// TwinCAT 3 PLC project IAG50cmTests
// Title: IAG50cmTests
// Company: BROT
// ProjectVersion: 0.1.0
// ProgramVersion: 3.1.4024.66
// libraries:
//   AstroBROT, 0.5.0 (BROT)
//   BROTLib, 0.20.0 (BROT)
//   Tc2_Math, * (Beckhoff Automation GmbH)
//   Tc3_MC2_AdvancedHoming, * (Beckhoff Automation GmbH)
//   Tc2_MC2, * (Beckhoff Automation GmbH)
//   Tc2_MC2_Drive, * (Beckhoff Automation GmbH)
//   Tc2_NC, * (Beckhoff Automation GmbH)
//   Tc2_Standard, * (Beckhoff Automation GmbH)
//   Tc2_System, * (Beckhoff Automation GmbH)
//   Tc2_Utilities, * (Beckhoff Automation GmbH)
//   Tc3_Module, * (Beckhoff Automation GmbH)
//   TcUnit, * (www.tcunit.org)
// project tree:
//   / PlcTask.TcTTO
//   POUs/ FB_HomeDropReason_Tests.TcPOU, FB_HomeHold_Tests.TcPOU, FB_SweepStop_Tests.TcPOU, FB_PointingModelForward_Tests.TcPOU, FB_TelescopeControl.TcPOU (not stored), FB_HourAngleControl.TcPOU (not stored), FB_DeclinationControl.TcPOU (not stored), FB_AxisControl.TcPOU (not stored), FB_LatchHome.TcPOU (not stored), FB_CabinetControl.TcPOU (not stored), FB_PointingModelInversion.TcPOU (not stored), F_HourAngleOffsetOnAxis.TcPOU (not stored), F_RoundLREAL.TcPOU (not stored), NCError_TO_STRING.TcPOU (not stored), ST_AxisStatus.TcDUT (not stored), FB_AxisMockCore.TcPOU, FB_HourAngleMock.TcPOU, FB_DeclinationMock.TcPOU, FB_FocusMock.TcPOU, FB_CoversMock.TcPOU, FB_DomeMock.TcPOU, FB_NullComm.TcPOU, FB_IagRig_Tests.TcPOU, FB_IagRig.TcPOU, IagStopDuringSlew_Tests.TcPOU, IagCommandInputs_Tests.TcPOU, IagCommandAcceptance_Tests.TcPOU, IagAbortStop_Tests.TcPOU, IagParkPowerReset_Tests.TcPOU, IagSupersede_Tests.TcPOU, IagStuckStop_Tests.TcPOU, GVL_Diag.TcGVL, F_Note.TcPOU, IagResetUnderMotion_Tests.TcPOU, IagTimeouts_Tests.TcPOU, IagErrorPark_Tests.TcPOU, IagParkDuringPowerOn_Tests.TcPOU, IagStopDuringPark_Tests.TcPOU, IagParkInLimit_Tests.TcPOU, FB_RecordingComm.TcPOU, F_NoteNear.TcPOU, FB_IagCoordinatesLegacy.TcPOU, IagTelemetry_Tests.TcPOU, IagCoordinates_Tests.TcPOU, MAIN.TcPOU, FB_HomeDropReason.TcPOU (not stored), FB_HomeHold.TcPOU (not stored), FB_StartRequest.TcPOU (not stored), FB_StartRequest_Tests.TcPOU, FB_StepDrain.TcPOU (not stored), FB_StepDrain_Tests.TcPOU, FB_SweepStop.TcPOU (not stored), FB_PointingModelForward.TcPOU (not stored), GVL_Homing.TcGVL (not stored), GVL_Pointing.TcGVL (not stored)
// real-time tasks:
//   TASK PlcTask: cycle T#10ms, priority 20, ADS port 350

CONFIGURATION IAG50cmTests
    RESOURCE PLC ON TwinCAT3
        TASK PlcTask(INTERVAL := T#10ms, PRIORITY := 20);
        PROGRAM MAIN WITH PlcTask : MAIN;
    END_RESOURCE
END_CONFIGURATION

// ---- POUs/GVL_Diag.TcGVL
{attribute 'qualified_only'}
VAR_GLOBAL
	// the failed checks of the scenario tests (F_Note), one "test: message;" each. Run-Tests.ps1 prints it when a test failed:
	// TcUnit itself only writes the failure text to the ADS log, which CI cannot see.
	sFailures	: STRING(1000);
END_VAR

// ---- POUs/MAIN.TcPOU
PROGRAM MAIN
VAR
	// TcUnit finds every FB_TestSuite instance by itself; it is enough to declare them here.
	fbHomeDropReasonTests	: FB_HomeDropReason_Tests;
	fbHomeHoldTests			: FB_HomeHold_Tests;
	fbStartRequestTests		: FB_StartRequest_Tests;
	fbStepDrainTests		: FB_StepDrain_Tests;
	fbSweepStopTests		: FB_SweepStop_Tests;
	fbPointingForwardTests	: FB_PointingModelForward_Tests;
	fbIagRigTests			: FB_IagRig_Tests;
	fbStopDuringSlewTests	: IagStopDuringSlew_Tests;
	fbResetUnderMotionTests	: IagResetUnderMotion_Tests;
	fbErrorParkTests		: IagErrorPark_Tests;
	fbIagTimeoutsTests : IagTimeouts_Tests;
	fbParkDuringPowerOnTests	: IagParkDuringPowerOn_Tests;
	fbStopDuringParkTests	: IagStopDuringPark_Tests;
	fbParkInLimitTests		: IagParkInLimit_Tests;
	fbStuckStopTests		: IagStuckStop_Tests;
	fbCommandInputsTests	: IagCommandInputs_Tests;
	fbCommandAcceptanceTests	: IagCommandAcceptance_Tests;
	fbAbortStopTests		: IagAbortStop_Tests;
	fbParkPowerResetTests	: IagParkPowerReset_Tests;
	fbSupersedeTests		: IagSupersede_Tests;
	fbTelemetryTests		: IagTelemetry_Tests;
	fbCoordinatesTests		: IagCoordinates_Tests;
END_VAR

TcUnit.RUN();

END_PROGRAM

// ---- POUs/FB_HomeDropReason_Tests.TcPOU
// Tests for FB_HomeDropReason, the text of the WARN when a pending home is dropped after 2 min (#108, #120).
FUNCTION_BLOCK FB_HomeDropReason_Tests EXTENDS TcUnit.FB_TestSuite
VAR
END_VAR

Not_Ready();
Stop_Did_Not_Finish();
Axes_Busy();
Not_Ready_Wins_Over_Stop_Pending();
Texts_Fit_Their_Strings();

METHOD PRIVATE Not_Ready
VAR
	fbHome	: FB_HomeDropReason;
END_VAR
TEST('Not_Ready');
fbHome(bReady := FALSE, bStopPending := FALSE);
AssertEquals_STRING(Expected := 'cancelled: telescope not ready', Actual := fbHome.sEnd, Message := 'sEnd');
AssertEquals_STRING(Expected := 'the telescope was not ready for 2 min. Power on, then send the home again.', Actual := fbHome.sWhy, Message := 'sWhy');
TEST_FINISHED();
END_METHOD

METHOD PRIVATE Stop_Did_Not_Finish
VAR
	fbHome	: FB_HomeDropReason;
END_VAR
TEST('Stop_Did_Not_Finish');
fbHome(bReady := TRUE, bStopPending := TRUE);
AssertEquals_STRING(Expected := 'cancelled: stop did not finish', Actual := fbHome.sEnd, Message := 'sEnd');
AssertEquals_STRING(Expected := 'the stop before the home did not finish within 2 min. Send the stop, then the home again.', Actual := fbHome.sWhy, Message := 'sWhy');
TEST_FINISHED();
END_METHOD

METHOD PRIVATE Axes_Busy
VAR
	fbHome	: FB_HomeDropReason;
END_VAR
TEST('Axes_Busy');
fbHome(bReady := TRUE, bStopPending := FALSE);
AssertEquals_STRING(Expected := 'cancelled: axes busy', Actual := fbHome.sEnd, Message := 'sEnd');
AssertEquals_STRING(Expected := 'the axes were busy for 2 min. Send the home again.', Actual := fbHome.sWhy, Message := 'sWhy');
TEST_FINISHED();
END_METHOD

METHOD PRIVATE Not_Ready_Wins_Over_Stop_Pending
VAR
	fbHome	: FB_HomeDropReason;
END_VAR
TEST('Not_Ready_Wins_Over_Stop_Pending');
fbHome(bReady := FALSE, bStopPending := TRUE);
AssertEquals_STRING(Expected := 'cancelled: telescope not ready', Actual := fbHome.sEnd, Message := 'sEnd');
AssertEquals_STRING(Expected := 'the telescope was not ready for 2 min. Power on, then send the home again.', Actual := fbHome.sWhy, Message := 'sWhy');
TEST_FINISHED();
END_METHOD

METHOD PRIVATE Texts_Fit_Their_Strings
VAR
	fbHome	: FB_HomeDropReason;
END_VAR
TEST('Texts_Fit_Their_Strings');
fbHome(bReady := TRUE, bStopPending := TRUE);
AssertEquals_BOOL(Expected := TRUE, Actual := LEN(fbHome.sEnd) < 40, Message := 'sEnd not cut off');
AssertEquals_BOOL(Expected := TRUE, Actual := LEN(fbHome.sWhy) < 160, Message := 'sWhy not cut off');
TEST_FINISHED();
END_METHOD

END_FUNCTION_BLOCK

// ---- POUs/FB_HomeHold_Tests.TcPOU
// Tests for FB_HomeHold, the no-new-homing-request after a stop in the calibration sweep (#113).
FUNCTION_BLOCK FB_HomeHold_Tests EXTENDS TcUnit.FB_TestSuite
VAR
END_VAR

No_Hold_Without_Stop();
Stop_While_Homing_Holds();
Hold_Stays_After_Stop_Done();
Stop_While_Not_Homing_Does_Not_Hold();
Stop_While_Calibrated_Does_Not_Hold();
Disable_Releases_The_Hold();
Reset_Releases_The_Hold();
New_PowerOn_Releases_The_Hold();
Release_Ignored_While_Stop_Active();
Release_Without_Hold_Changes_Nothing();
StopSweep_Holds_An_Uncalibrated_Axis_Before_The_Sweep_Starts();
StopSweep_Ignored_On_A_Calibrated_Axis();
StopSweep_Wins_Over_Release_In_The_Same_Scan();
StopSweep_Hold_Ends_With_Disable();
StopSweep_Hold_Ends_With_Release_In_A_Later_Scan();

METHOD PRIVATE No_Hold_Without_Stop
VAR
	fbHold	: FB_HomeHold;
END_VAR
TEST('No_Hold_Without_Stop');
fbHold(bEnable := TRUE, bCalibrated := FALSE, bHoming := TRUE, bStopAxis := FALSE, bReset := FALSE);
AssertEquals_BOOL(Expected := FALSE, Actual := fbHold.bHold, Message := 'homing runs');
TEST_FINISHED();
END_METHOD

METHOD PRIVATE Stop_While_Homing_Holds
VAR
	fbHold	: FB_HomeHold;
END_VAR
TEST('Stop_While_Homing_Holds');
fbHold(bEnable := TRUE, bCalibrated := FALSE, bHoming := TRUE, bStopAxis := FALSE, bReset := FALSE);
fbHold(bEnable := TRUE, bCalibrated := FALSE, bHoming := TRUE, bStopAxis := TRUE, bReset := FALSE);
AssertEquals_BOOL(Expected := TRUE, Actual := fbHold.bHold, Message := 'held after the stop');
TEST_FINISHED();
END_METHOD

METHOD PRIVATE Hold_Stays_After_Stop_Done
VAR
	fbHold	: FB_HomeHold;
END_VAR
TEST('Hold_Stays_After_Stop_Done');
// bStopAxis falls on StopDone, bHomeAxis is cleared by the hold: the hold must stay while the axis is enabled
fbHold(bEnable := TRUE, bCalibrated := FALSE, bHoming := TRUE, bStopAxis := FALSE, bReset := FALSE);
fbHold(bEnable := TRUE, bCalibrated := FALSE, bHoming := TRUE, bStopAxis := TRUE, bReset := FALSE);
fbHold(bEnable := TRUE, bCalibrated := FALSE, bHoming := FALSE, bStopAxis := FALSE, bReset := FALSE);
fbHold(bEnable := TRUE, bCalibrated := FALSE, bHoming := FALSE, bStopAxis := FALSE, bReset := FALSE);
AssertEquals_BOOL(Expected := TRUE, Actual := fbHold.bHold, Message := 'still held');
TEST_FINISHED();
END_METHOD

METHOD PRIVATE Stop_While_Not_Homing_Does_Not_Hold
VAR
	fbHold	: FB_HomeHold;
END_VAR
TEST('Stop_While_Not_Homing_Does_Not_Hold');
fbHold(bEnable := TRUE, bCalibrated := FALSE, bHoming := FALSE, bStopAxis := TRUE, bReset := FALSE);
AssertEquals_BOOL(Expected := FALSE, Actual := fbHold.bHold, Message := 'no sweep, no hold');
TEST_FINISHED();
END_METHOD

METHOD PRIVATE Stop_While_Calibrated_Does_Not_Hold
VAR
	fbHold	: FB_HomeHold;
END_VAR
TEST('Stop_While_Calibrated_Does_Not_Hold');
fbHold(bEnable := TRUE, bCalibrated := TRUE, bHoming := TRUE, bStopAxis := TRUE, bReset := FALSE);
AssertEquals_BOOL(Expected := FALSE, Actual := fbHold.bHold, Message := 'calibrated');
TEST_FINISHED();
END_METHOD

METHOD PRIVATE Disable_Releases_The_Hold
VAR
	fbHold	: FB_HomeHold;
END_VAR
TEST('Disable_Releases_The_Hold');
fbHold(bEnable := TRUE, bCalibrated := FALSE, bHoming := TRUE, bStopAxis := FALSE, bReset := FALSE);
fbHold(bEnable := TRUE, bCalibrated := FALSE, bHoming := TRUE, bStopAxis := TRUE, bReset := FALSE);
fbHold(bEnable := FALSE, bCalibrated := FALSE, bHoming := FALSE, bStopAxis := FALSE, bReset := FALSE);
AssertEquals_BOOL(Expected := FALSE, Actual := fbHold.bHold, Message := 'released');
fbHold(bEnable := TRUE, bCalibrated := FALSE, bHoming := TRUE, bStopAxis := FALSE, bReset := FALSE);
AssertEquals_BOOL(Expected := FALSE, Actual := fbHold.bHold, Message := 'homing again');
TEST_FINISHED();
END_METHOD

METHOD PRIVATE Reset_Releases_The_Hold
VAR
	fbHold	: FB_HomeHold;
END_VAR
TEST('Reset_Releases_The_Hold');
fbHold(bEnable := TRUE, bCalibrated := FALSE, bHoming := TRUE, bStopAxis := FALSE, bReset := FALSE);
fbHold(bEnable := TRUE, bCalibrated := FALSE, bHoming := TRUE, bStopAxis := TRUE, bReset := FALSE);
fbHold(bEnable := TRUE, bCalibrated := FALSE, bHoming := FALSE, bStopAxis := FALSE, bReset := TRUE);
AssertEquals_BOOL(Expected := FALSE, Actual := fbHold.bHold, Message := 'released by reset');
TEST_FINISHED();
END_METHOD

METHOD PRIVATE New_PowerOn_Releases_The_Hold
VAR
	fbHold	: FB_HomeHold;
END_VAR
TEST('New_PowerOn_Releases_The_Hold');
// an automatic stop at stage 40: held, axis still enabled, reset=1 gives no bReset (#159)
fbHold(bEnable := TRUE, bCalibrated := FALSE, bHoming := TRUE, bStopAxis := FALSE, bReset := FALSE);
fbHold(bEnable := TRUE, bCalibrated := FALSE, bHoming := TRUE, bStopAxis := TRUE, bReset := FALSE);
fbHold(bEnable := TRUE, bCalibrated := FALSE, bHoming := FALSE, bStopAxis := FALSE, bReset := FALSE);
AssertEquals_BOOL(Expected := TRUE, Actual := fbHold.bHold, Message := 'held');
fbHold(bEnable := TRUE, bCalibrated := FALSE, bHoming := FALSE, bStopAxis := FALSE, bReset := FALSE, bRelease := TRUE);
AssertEquals_BOOL(Expected := FALSE, Actual := fbHold.bHold, Message := 'released by the new power-on');
TEST_FINISHED();
END_METHOD

METHOD PRIVATE Release_Ignored_While_Stop_Active
VAR
	fbHold	: FB_HomeHold;
END_VAR
TEST('Release_Ignored_While_Stop_Active');
fbHold(bEnable := TRUE, bCalibrated := FALSE, bHoming := TRUE, bStopAxis := FALSE, bReset := FALSE);
fbHold(bEnable := TRUE, bCalibrated := FALSE, bHoming := TRUE, bStopAxis := TRUE, bReset := FALSE, bRelease := TRUE);
AssertEquals_BOOL(Expected := TRUE, Actual := fbHold.bHold, Message := 'a running stop is not cut through');
TEST_FINISHED();
END_METHOD

METHOD PRIVATE Release_Without_Hold_Changes_Nothing
VAR
	fbHold	: FB_HomeHold;
END_VAR
TEST('Release_Without_Hold_Changes_Nothing');
fbHold(bEnable := TRUE, bCalibrated := FALSE, bHoming := TRUE, bStopAxis := FALSE, bReset := FALSE, bRelease := TRUE);
AssertEquals_BOOL(Expected := FALSE, Actual := fbHold.bHold, Message := 'no hold');
TEST_FINISHED();
END_METHOD

METHOD PRIVATE StopSweep_Holds_An_Uncalibrated_Axis_Before_The_Sweep_Starts
VAR
	fbHold	: FB_HomeHold;
END_VAR
TEST('StopSweep_Holds_An_Uncalibrated_Axis_Before_The_Sweep_Starts');
// #198: the stop arrives before bHomeAxis is set (tonReady, or the scans after a reset)
fbHold(bEnable := TRUE, bCalibrated := FALSE, bHoming := FALSE, bStopAxis := FALSE, bReset := FALSE, bStopSweep := TRUE);
AssertEquals_BOOL(Expected := TRUE, Actual := fbHold.bHold, Message := 'held');
fbHold(bEnable := TRUE, bCalibrated := FALSE, bHoming := FALSE, bStopAxis := FALSE, bReset := FALSE, bStopSweep := FALSE);
AssertEquals_BOOL(Expected := TRUE, Actual := fbHold.bHold, Message := 'still held');
TEST_FINISHED();
END_METHOD

METHOD PRIVATE StopSweep_Ignored_On_A_Calibrated_Axis
VAR
	fbHold	: FB_HomeHold;
END_VAR
TEST('StopSweep_Ignored_On_A_Calibrated_Axis');
fbHold(bEnable := TRUE, bCalibrated := TRUE, bHoming := FALSE, bStopAxis := FALSE, bReset := FALSE, bStopSweep := TRUE);
AssertEquals_BOOL(Expected := FALSE, Actual := fbHold.bHold, Message := 'calibrated axis not held');
TEST_FINISHED();
END_METHOD

METHOD PRIVATE StopSweep_Wins_Over_Release_In_The_Same_Scan
VAR
	fbHold	: FB_HomeHold;
END_VAR
TEST('StopSweep_Wins_Over_Release_In_The_Same_Scan');
fbHold(bEnable := TRUE, bCalibrated := FALSE, bHoming := FALSE, bStopAxis := FALSE, bReset := FALSE, bRelease := TRUE, bStopSweep := TRUE);
AssertEquals_BOOL(Expected := TRUE, Actual := fbHold.bHold, Message := 'held');
TEST_FINISHED();
END_METHOD

METHOD PRIVATE StopSweep_Hold_Ends_With_Disable
VAR
	fbHold	: FB_HomeHold;
END_VAR
TEST('StopSweep_Hold_Ends_With_Disable');
fbHold(bEnable := TRUE, bCalibrated := FALSE, bHoming := FALSE, bStopAxis := FALSE, bReset := FALSE, bStopSweep := TRUE);
fbHold(bEnable := FALSE, bCalibrated := FALSE, bHoming := FALSE, bStopAxis := FALSE, bReset := FALSE, bStopSweep := FALSE);
AssertEquals_BOOL(Expected := FALSE, Actual := fbHold.bHold, Message := 'released by the disable');
TEST_FINISHED();
END_METHOD

METHOD PRIVATE StopSweep_Hold_Ends_With_Release_In_A_Later_Scan
VAR
	fbHold	: FB_HomeHold;
END_VAR
TEST('StopSweep_Hold_Ends_With_Release_In_A_Later_Scan');
fbHold(bEnable := TRUE, bCalibrated := FALSE, bHoming := FALSE, bStopAxis := FALSE, bReset := FALSE, bStopSweep := TRUE);
fbHold(bEnable := TRUE, bCalibrated := FALSE, bHoming := FALSE, bStopAxis := FALSE, bReset := FALSE, bRelease := TRUE, bStopSweep := FALSE);
AssertEquals_BOOL(Expected := FALSE, Actual := fbHold.bHold, Message := 'released by a new power-on');
TEST_FINISHED();
END_METHOD

END_FUNCTION_BLOCK

// ---- POUs/FB_StartRequest_Tests.TcPOU
// Tests for FB_StartRequest, the start request of FB_LatchHome that must survive an abort in progress (#155).
FUNCTION_BLOCK FB_StartRequest_Tests EXTENDS TcUnit.FB_TestSuite
VAR
END_VAR

Edge_Is_Taken_Once();
Edge_While_Busy_Is_Kept();
No_Restart_While_Execute_Stays_True();
Execute_Falling_Drops_The_Request();
New_Edge_Starts_Again();
Rearm_Asks_Again_While_Execute_Is_True();
Rearm_Does_Nothing_Without_Execute();
Pending_Survives_Until_Taken_Later();

METHOD PRIVATE Edge_Is_Taken_Once
VAR
	fbReq	: FB_StartRequest;
END_VAR
TEST('Edge_Is_Taken_Once');
fbReq(Execute := FALSE);
fbReq(Execute := TRUE);
AssertEquals_BOOL(Expected := TRUE, Actual := fbReq.Take(), Message := 'first take');
AssertEquals_BOOL(Expected := FALSE, Actual := fbReq.Take(), Message := 'second take');
TEST_FINISHED();
END_METHOD

METHOD PRIVATE Edge_While_Busy_Is_Kept
VAR
	fbReq	: FB_StartRequest;
	i		: INT;
END_VAR
TEST('Edge_While_Busy_Is_Kept');
// the edge arrives while the block is aborting and nobody takes it for a number of scans (#155)
fbReq(Execute := FALSE);
fbReq(Execute := TRUE);
FOR i := 1 TO 20 DO
	fbReq(Execute := TRUE);
END_FOR
AssertEquals_BOOL(Expected := TRUE, Actual := fbReq.Take(), Message := 'taken once the abort is over');
TEST_FINISHED();
END_METHOD

METHOD PRIVATE No_Restart_While_Execute_Stays_True
VAR
	fbReq	: FB_StartRequest;
END_VAR
TEST('No_Restart_While_Execute_Stays_True');
fbReq(Execute := FALSE);
fbReq(Execute := TRUE);
fbReq.Take();
fbReq(Execute := TRUE);
fbReq(Execute := TRUE);
AssertEquals_BOOL(Expected := FALSE, Actual := fbReq.Take(), Message := 'no new edge, no new start');
TEST_FINISHED();
END_METHOD

METHOD PRIVATE Execute_Falling_Drops_The_Request
VAR
	fbReq	: FB_StartRequest;
END_VAR
TEST('Execute_Falling_Drops_The_Request');
fbReq(Execute := FALSE);
fbReq(Execute := TRUE);
fbReq(Execute := FALSE);
AssertEquals_BOOL(Expected := FALSE, Actual := fbReq.Take(), Message := 'request withdrawn');
TEST_FINISHED();
END_METHOD

METHOD PRIVATE New_Edge_Starts_Again
VAR
	fbReq	: FB_StartRequest;
END_VAR
TEST('New_Edge_Starts_Again');
fbReq(Execute := FALSE);
fbReq(Execute := TRUE);
fbReq.Take();
fbReq(Execute := FALSE);
fbReq(Execute := TRUE);
AssertEquals_BOOL(Expected := TRUE, Actual := fbReq.Take(), Message := 'second sweep');
TEST_FINISHED();
END_METHOD

METHOD PRIVATE Rearm_Asks_Again_While_Execute_Is_True
VAR
	fbReq	: FB_StartRequest;
END_VAR
TEST('Rearm_Asks_Again_While_Execute_Is_True');
// the start was taken, ended in the abort state without a result and Execute stayed TRUE (#155)
fbReq(Execute := FALSE);
fbReq(Execute := TRUE);
fbReq.Take();
fbReq(Execute := TRUE);
fbReq.Rearm();
AssertEquals_BOOL(Expected := TRUE, Actual := fbReq.Take(), Message := 'started again');
AssertEquals_BOOL(Expected := FALSE, Actual := fbReq.Take(), Message := 'once');
TEST_FINISHED();
END_METHOD

METHOD PRIVATE Rearm_Does_Nothing_Without_Execute
VAR
	fbReq	: FB_StartRequest;
END_VAR
TEST('Rearm_Does_Nothing_Without_Execute');
fbReq(Execute := FALSE);
fbReq.Rearm();
AssertEquals_BOOL(Expected := FALSE, Actual := fbReq.Take(), Message := 'no request');
TEST_FINISHED();
END_METHOD

METHOD PRIVATE Pending_Survives_Until_Taken_Later
VAR
	fbReq	: FB_StartRequest;
	i		: INT;
END_VAR
TEST('Pending_Survives_Until_Taken_Later');
// FB_LatchHome takes no start while a step block is still Busy (#113): the request must wait for it
fbReq(Execute := FALSE);
fbReq(Execute := TRUE);
FOR i := 1 TO 50 DO
	fbReq(Execute := TRUE);
END_FOR
AssertEquals_BOOL(Expected := TRUE, Actual := fbReq.Pending, Message := 'still pending');
AssertEquals_BOOL(Expected := TRUE, Actual := fbReq.Take(), Message := 'taken later');
AssertEquals_BOOL(Expected := FALSE, Actual := fbReq.Take(), Message := 'once');
TEST_FINISHED();
END_METHOD

END_FUNCTION_BLOCK

// ---- POUs/FB_StepDrain_Tests.TcPOU
// Tests for FB_StepDrain, the drain of a stale step block before FB_LatchHome takes a start (#113).
FUNCTION_BLOCK FB_StepDrain_Tests EXTENDS TcUnit.FB_TestSuite
VAR
END_VAR

Idle_Not_Busy_May_Take();
Busy_Drains_And_Blocks_Start();
No_Drain_Outside_Idle();
Start_Taken_Once_Busy_Drops();
Stuck_Only_With_Pending_Start();
Busy_Dropping_Before_Timeout_Is_Not_Stuck();

METHOD PRIVATE Idle_Not_Busy_May_Take
VAR
	fbDrain	: FB_StepDrain;
END_VAR
TEST('Idle_Not_Busy_May_Take');
fbDrain(bIdle := TRUE, bStepBusy := FALSE, bStartPending := TRUE);
AssertEquals_BOOL(Expected := TRUE, Actual := fbDrain.bMayTake, Message := 'may take');
AssertEquals_BOOL(Expected := FALSE, Actual := fbDrain.bDrain, Message := 'no drain');
TEST_FINISHED();
END_METHOD

METHOD PRIVATE Busy_Drains_And_Blocks_Start
VAR
	fbDrain	: FB_StepDrain;
END_VAR
TEST('Busy_Drains_And_Blocks_Start');
fbDrain(bIdle := TRUE, bStepBusy := TRUE, bStartPending := TRUE, PT := T#1H);
AssertEquals_BOOL(Expected := TRUE, Actual := fbDrain.bDrain, Message := 'drain');
AssertEquals_BOOL(Expected := FALSE, Actual := fbDrain.bMayTake, Message := 'no start while busy');
AssertEquals_BOOL(Expected := FALSE, Actual := fbDrain.bStuck, Message := 'not stuck yet');
TEST_FINISHED();
END_METHOD

METHOD PRIVATE No_Drain_Outside_Idle
VAR
	fbDrain	: FB_StepDrain;
END_VAR
TEST('No_Drain_Outside_Idle');
fbDrain(bIdle := FALSE, bStepBusy := TRUE, bStartPending := TRUE, PT := T#0S);
AssertEquals_BOOL(Expected := FALSE, Actual := fbDrain.bDrain, Message := 'a running step is not released');
AssertEquals_BOOL(Expected := FALSE, Actual := fbDrain.bMayTake, Message := 'no start outside idle');
AssertEquals_BOOL(Expected := FALSE, Actual := fbDrain.bStuck, Message := 'not stuck outside idle');
TEST_FINISHED();
END_METHOD

METHOD PRIVATE Start_Taken_Once_Busy_Drops
VAR
	fbDrain	: FB_StepDrain;
	fbReq	: FB_StartRequest;
	i		: INT;
	nTaken	: INT;
END_VAR
TEST('Start_Taken_Once_Busy_Drops');
// the sequence of the 14:07 run: a start waits while the stale block drains, then it is taken exactly once
fbReq(Execute := FALSE);
fbReq(Execute := TRUE);
FOR i := 1 TO 5 DO
	fbDrain(bIdle := TRUE, bStepBusy := TRUE, bStartPending := fbReq.Pending, PT := T#1H);
	// nested like FB_LatchHome: AND does not short-circuit, Take() would clear the pending request while the block is busy
	IF fbDrain.bMayTake THEN
		IF fbReq.Take() THEN
			nTaken := nTaken + 1;
		END_IF
	END_IF
END_FOR
AssertEquals_INT(Expected := 0, Actual := nTaken, Message := 'nothing taken while busy');
FOR i := 1 TO 5 DO
	fbReq(Execute := TRUE);
	fbDrain(bIdle := TRUE, bStepBusy := FALSE, bStartPending := fbReq.Pending, PT := T#1H);
	// nested like FB_LatchHome: AND does not short-circuit, Take() would clear the pending request while the block is busy
	IF fbDrain.bMayTake THEN
		IF fbReq.Take() THEN
			nTaken := nTaken + 1;
		END_IF
	END_IF
END_FOR
AssertEquals_INT(Expected := 1, Actual := nTaken, Message := 'taken once after the drain');
TEST_FINISHED();
END_METHOD

METHOD PRIVATE Stuck_Only_With_Pending_Start
VAR
	fbDrain	: FB_StepDrain;
END_VAR
TEST('Stuck_Only_With_Pending_Start');
fbDrain(bIdle := TRUE, bStepBusy := TRUE, bStartPending := FALSE, PT := T#0S);
AssertEquals_BOOL(Expected := FALSE, Actual := fbDrain.bStuck, Message := 'a busy block without a start is no error');
fbDrain(bIdle := TRUE, bStepBusy := TRUE, bStartPending := TRUE, PT := T#0S);
AssertEquals_BOOL(Expected := TRUE, Actual := fbDrain.bStuck, Message := 'stuck with a pending start');
TEST_FINISHED();
END_METHOD

METHOD PRIVATE Busy_Dropping_Before_Timeout_Is_Not_Stuck
VAR
	fbDrain	: FB_StepDrain;
END_VAR
TEST('Busy_Dropping_Before_Timeout_Is_Not_Stuck');
fbDrain(bIdle := TRUE, bStepBusy := TRUE, bStartPending := TRUE, PT := T#1H);
fbDrain(bIdle := TRUE, bStepBusy := FALSE, bStartPending := TRUE, PT := T#1H);
AssertEquals_BOOL(Expected := FALSE, Actual := fbDrain.bStuck, Message := 'not stuck');
AssertEquals_BOOL(Expected := TRUE, Actual := fbDrain.bMayTake, Message := 'may take');
TEST_FINISHED();
END_METHOD

END_FUNCTION_BLOCK

// ---- POUs/FB_SweepStop_Tests.TcPOU
// Tests for FB_SweepStop, switching the uncalibrated axes off after a stop in the calibration sweep (#113).
FUNCTION_BLOCK FB_SweepStop_Tests EXTENDS TcUnit.FB_TestSuite
VAR
END_VAR

Disables_Uncalibrated_Axes_After_Three_Settled_Scans();
Calibrated_Axis_Stays_Enabled();
Waits_While_Homing_Runs();
Not_Settled_Restarts_The_Count();
No_Disable_Without_Arm();
Disable_Is_A_One_Scan_Pulse();
Cancel_Drops_The_Request();
ArmAll_Disables_Calibrated_Axes_Too();
ArmAll_Is_Idempotent();
ArmAll_Waits_For_The_Focus();
Arm_Ignores_OtherBusy();
Arm_Does_Not_Narrow_A_Pending_ArmAll();
Cancel_Clears_All_Mode();

METHOD PRIVATE Disables_Uncalibrated_Axes_After_Three_Settled_Scans
VAR
	fbSw	: FB_SweepStop;
	i		: INT;
END_VAR
TEST('Disables_Uncalibrated_Axes_After_Three_Settled_Scans');
fbSw.Arm();
FOR i := 1 TO 2 DO
fbSw(bSettled := TRUE, bHaCalibrated := FALSE, bDecCalibrated := FALSE, bHaHoming := FALSE, bDecHoming := FALSE);
END_FOR
AssertEquals_BOOL(Expected := FALSE, Actual := fbSw.bDisableHa, Message := 'two scans: not yet');
fbSw(bSettled := TRUE, bHaCalibrated := FALSE, bDecCalibrated := FALSE, bHaHoming := FALSE, bDecHoming := FALSE);
AssertEquals_BOOL(Expected := TRUE, Actual := fbSw.bDisableHa, Message := 'HA off');
AssertEquals_BOOL(Expected := TRUE, Actual := fbSw.bDisableDec, Message := 'Dec off');
TEST_FINISHED();
END_METHOD

METHOD PRIVATE Calibrated_Axis_Stays_Enabled
VAR
	fbSw	: FB_SweepStop;
	i		: INT;
END_VAR
TEST('Calibrated_Axis_Stays_Enabled');
fbSw.Arm();
FOR i := 1 TO 3 DO
fbSw(bSettled := TRUE, bHaCalibrated := TRUE, bDecCalibrated := FALSE, bHaHoming := FALSE, bDecHoming := FALSE);
END_FOR
AssertEquals_BOOL(Expected := FALSE, Actual := fbSw.bDisableHa, Message := 'HA calibrated');
AssertEquals_BOOL(Expected := TRUE, Actual := fbSw.bDisableDec, Message := 'Dec off');
TEST_FINISHED();
END_METHOD

METHOD PRIVATE Waits_While_Homing_Runs
VAR
	fbSw	: FB_SweepStop;
	i		: INT;
END_VAR
TEST('Waits_While_Homing_Runs');
fbSw.Arm();
FOR i := 1 TO 50 DO
fbSw(bSettled := TRUE, bHaCalibrated := FALSE, bDecCalibrated := FALSE, bHaHoming := TRUE, bDecHoming := FALSE);
END_FOR
AssertEquals_BOOL(Expected := FALSE, Actual := fbSw.bDisableHa, Message := 'HA homing busy');
FOR i := 1 TO 50 DO
fbSw(bSettled := TRUE, bHaCalibrated := FALSE, bDecCalibrated := FALSE, bHaHoming := FALSE, bDecHoming := TRUE);
END_FOR
AssertEquals_BOOL(Expected := FALSE, Actual := fbSw.bDisableDec, Message := 'Dec homing busy');
FOR i := 1 TO 3 DO
fbSw(bSettled := TRUE, bHaCalibrated := FALSE, bDecCalibrated := FALSE, bHaHoming := FALSE, bDecHoming := FALSE);
END_FOR
AssertEquals_BOOL(Expected := TRUE, Actual := fbSw.bDisableHa, Message := 'off when the homing is idle');
TEST_FINISHED();
END_METHOD

METHOD PRIVATE Not_Settled_Restarts_The_Count
VAR
	fbSw	: FB_SweepStop;
	i		: INT;
END_VAR
TEST('Not_Settled_Restarts_The_Count');
fbSw.Arm();
FOR i := 1 TO 2 DO
fbSw(bSettled := TRUE, bHaCalibrated := FALSE, bDecCalibrated := FALSE, bHaHoming := FALSE, bDecHoming := FALSE);
END_FOR
fbSw(bSettled := FALSE, bHaCalibrated := FALSE, bDecCalibrated := FALSE, bHaHoming := FALSE, bDecHoming := FALSE);
FOR i := 1 TO 2 DO
fbSw(bSettled := TRUE, bHaCalibrated := FALSE, bDecCalibrated := FALSE, bHaHoming := FALSE, bDecHoming := FALSE);
END_FOR
AssertEquals_BOOL(Expected := FALSE, Actual := fbSw.bDisableHa, Message := 'count restarted');
fbSw(bSettled := TRUE, bHaCalibrated := FALSE, bDecCalibrated := FALSE, bHaHoming := FALSE, bDecHoming := FALSE);
AssertEquals_BOOL(Expected := TRUE, Actual := fbSw.bDisableHa, Message := 'off');
TEST_FINISHED();
END_METHOD

METHOD PRIVATE No_Disable_Without_Arm
VAR
	fbSw	: FB_SweepStop;
	i		: INT;
END_VAR
TEST('No_Disable_Without_Arm');
FOR i := 1 TO 20 DO
fbSw(bSettled := TRUE, bHaCalibrated := FALSE, bDecCalibrated := FALSE, bHaHoming := FALSE, bDecHoming := FALSE);
END_FOR
AssertEquals_BOOL(Expected := FALSE, Actual := fbSw.bDisableHa, Message := 'not armed');
AssertEquals_BOOL(Expected := FALSE, Actual := fbSw.bDisableDec, Message := 'not armed');
TEST_FINISHED();
END_METHOD

METHOD PRIVATE Disable_Is_A_One_Scan_Pulse
VAR
	fbSw	: FB_SweepStop;
	i		: INT;
END_VAR
TEST('Disable_Is_A_One_Scan_Pulse');
fbSw.Arm();
FOR i := 1 TO 3 DO
fbSw(bSettled := TRUE, bHaCalibrated := FALSE, bDecCalibrated := FALSE, bHaHoming := FALSE, bDecHoming := FALSE);
END_FOR
AssertEquals_BOOL(Expected := TRUE, Actual := fbSw.bDisableHa, Message := 'pulse');
fbSw(bSettled := TRUE, bHaCalibrated := FALSE, bDecCalibrated := FALSE, bHaHoming := FALSE, bDecHoming := FALSE);
AssertEquals_BOOL(Expected := FALSE, Actual := fbSw.bDisableHa, Message := 'only once');
AssertEquals_BOOL(Expected := FALSE, Actual := fbSw.bDisableDec, Message := 'only once');
TEST_FINISHED();
END_METHOD

METHOD PRIVATE Cancel_Drops_The_Request
VAR
	fbSw	: FB_SweepStop;
	i		: INT;
END_VAR
TEST('Cancel_Drops_The_Request');
fbSw.Arm();
FOR i := 1 TO 2 DO
fbSw(bSettled := TRUE, bHaCalibrated := FALSE, bDecCalibrated := FALSE, bHaHoming := FALSE, bDecHoming := FALSE);
END_FOR
fbSw.Cancel();
FOR i := 1 TO 10 DO
fbSw(bSettled := TRUE, bHaCalibrated := FALSE, bDecCalibrated := FALSE, bHaHoming := FALSE, bDecHoming := FALSE);
END_FOR
AssertEquals_BOOL(Expected := FALSE, Actual := fbSw.bDisableHa, Message := 'cancelled');
TEST_FINISHED();
END_METHOD

// #197: a park without a completed power-on switches every axis off, calibrated or not
METHOD PRIVATE ArmAll_Disables_Calibrated_Axes_Too
VAR
	fbSw	: FB_SweepStop;
	i		: INT;
END_VAR
TEST('ArmAll_Disables_Calibrated_Axes_Too');
fbSw.ArmAll();
FOR i := 1 TO 2 DO
fbSw(bSettled := TRUE, bHaCalibrated := TRUE, bDecCalibrated := TRUE, bHaHoming := FALSE, bDecHoming := FALSE);
END_FOR
AssertEquals_BOOL(Expected := FALSE, Actual := fbSw.bDisableHa, Message := 'two scans: not yet');
fbSw(bSettled := TRUE, bHaCalibrated := TRUE, bDecCalibrated := TRUE, bHaHoming := FALSE, bDecHoming := FALSE);
AssertEquals_BOOL(Expected := TRUE, Actual := fbSw.bDisableHa, Message := 'HA off although calibrated');
AssertEquals_BOOL(Expected := TRUE, Actual := fbSw.bDisableDec, Message := 'Dec off although calibrated');
fbSw(bSettled := TRUE, bHaCalibrated := TRUE, bDecCalibrated := TRUE, bHaHoming := FALSE, bDecHoming := FALSE);
AssertEquals_BOOL(Expected := FALSE, Actual := fbSw.bDisableHa, Message := 'one scan only');
TEST_FINISHED();
END_METHOD

// #197: the arbitration calls ArmAll every scan
METHOD PRIVATE ArmAll_Is_Idempotent
VAR
	fbSw	: FB_SweepStop;
	i		: INT;
END_VAR
TEST('ArmAll_Is_Idempotent');
FOR i := 1 TO 2 DO
fbSw.ArmAll();
fbSw(bSettled := TRUE, bHaCalibrated := TRUE, bDecCalibrated := TRUE, bHaHoming := FALSE, bDecHoming := FALSE);
END_FOR
fbSw.ArmAll();
fbSw(bSettled := TRUE, bHaCalibrated := TRUE, bDecCalibrated := TRUE, bHaHoming := FALSE, bDecHoming := FALSE);
AssertEquals_BOOL(Expected := TRUE, Actual := fbSw.bDisableHa, Message := 'ArmAll every scan does not restart the count');
TEST_FINISHED();
END_METHOD

// #197: the focus must not be moving when the axes are switched off (#56)
METHOD PRIVATE ArmAll_Waits_For_The_Focus
VAR
	fbSw	: FB_SweepStop;
	i		: INT;
END_VAR
TEST('ArmAll_Waits_For_The_Focus');
fbSw.ArmAll();
FOR i := 1 TO 20 DO
fbSw(bSettled := TRUE, bHaCalibrated := TRUE, bDecCalibrated := TRUE, bHaHoming := FALSE, bDecHoming := FALSE, bOtherBusy := TRUE);
END_FOR
AssertEquals_BOOL(Expected := FALSE, Actual := fbSw.bDisableHa, Message := 'the focus is moving');
FOR i := 1 TO 3 DO
fbSw(bSettled := TRUE, bHaCalibrated := TRUE, bDecCalibrated := TRUE, bHaHoming := FALSE, bDecHoming := FALSE, bOtherBusy := FALSE);
END_FOR
AssertEquals_BOOL(Expected := TRUE, Actual := fbSw.bDisableDec, Message := 'off when the focus is at rest');
TEST_FINISHED();
END_METHOD

// #113 mode unchanged
METHOD PRIVATE Arm_Ignores_OtherBusy
VAR
	fbSw	: FB_SweepStop;
	i		: INT;
END_VAR
TEST('Arm_Ignores_OtherBusy');
fbSw.Arm();
FOR i := 1 TO 3 DO
fbSw(bSettled := TRUE, bHaCalibrated := FALSE, bDecCalibrated := TRUE, bHaHoming := FALSE, bDecHoming := FALSE, bOtherBusy := TRUE);
END_FOR
AssertEquals_BOOL(Expected := TRUE, Actual := fbSw.bDisableHa, Message := 'the stop of #113 does not wait for the focus');
AssertEquals_BOOL(Expected := FALSE, Actual := fbSw.bDisableDec, Message := 'calibrated axis stays on');
TEST_FINISHED();
END_METHOD

// a stop after the park request must not undo the all-axes mode
METHOD PRIVATE Arm_Does_Not_Narrow_A_Pending_ArmAll
VAR
	fbSw	: FB_SweepStop;
	i		: INT;
END_VAR
TEST('Arm_Does_Not_Narrow_A_Pending_ArmAll');
fbSw.ArmAll();
fbSw.Arm();
FOR i := 1 TO 3 DO
fbSw(bSettled := TRUE, bHaCalibrated := TRUE, bDecCalibrated := TRUE, bHaHoming := FALSE, bDecHoming := FALSE);
END_FOR
AssertEquals_BOOL(Expected := TRUE, Actual := fbSw.bDisableHa, Message := 'still the all-axes mode');
TEST_FINISHED();
END_METHOD

// Cancel drops the all-axes mode
METHOD PRIVATE Cancel_Clears_All_Mode
VAR
	fbSw	: FB_SweepStop;
	i		: INT;
END_VAR
TEST('Cancel_Clears_All_Mode');
fbSw.ArmAll();
fbSw.Cancel();
fbSw.Arm();
FOR i := 1 TO 3 DO
fbSw(bSettled := TRUE, bHaCalibrated := TRUE, bDecCalibrated := FALSE, bHaHoming := FALSE, bDecHoming := FALSE);
END_FOR
AssertEquals_BOOL(Expected := FALSE, Actual := fbSw.bDisableHa, Message := 'calibrated axis stays on after Cancel');
AssertEquals_BOOL(Expected := TRUE, Actual := fbSw.bDisableDec, Message := 'uncalibrated axis off');
TEST_FINISHED();
END_METHOD

END_FUNCTION_BLOCK

// ---- POUs/FB_PointingModelForward_Tests.TcPOU
// Tests for FB_PointingModelForward at the zenith (#4): finite outputs, continuity, unchanged values elsewhere.
FUNCTION_BLOCK FB_PointingModelForward_Tests EXTENDS TcUnit.FB_TestSuite
VAR
END_VAR

Zenith_Is_Finite();
Zenith_Velocity_Is_Sidereal();
Near_Zenith_Is_Continuous();
Reference_Points_Unchanged();

METHOD PRIVATE Zenith_Is_Finite
VAR
	fbModel	: FB_PointingModelForward;
	i		: INT;
	j		: INT;
	fLat	: LREAL;
	fHa		: LREAL;
	bOk		: BOOL := TRUE;
END_VAR
TEST('Zenith_Is_Finite');
// Dec = Lat, HA ~ 0, every latitude in 0.5 deg steps: sin_alt rounds to 1 + 2.2E-16 or exactly 1.0 for many of them (#4).
// ST has no ISNAN: ABS(x) < 1E3 is FALSE for NaN and Inf (the outputs are a few deg or deg/s at most)
FOR i := -179 TO 179 DO
	fLat := INT_TO_LREAL(i) * 0.5;
	FOR j := -1 TO 1 DO
		fHa := INT_TO_LREAL(j) * 1.0E-6;
		fbModel(HourAngle := fHa, Declination := fLat, Latitude := fLat);
		bOk := bOk AND (ABS(fbModel.HourAngle_correction) < 1.0E3) AND (ABS(fbModel.Declination_correction) < 1.0E3)
			AND (ABS(fbModel.HourAngle_velocity) < 1.0E3) AND (ABS(fbModel.Declination_velocity) < 1.0E3);
	END_FOR
END_FOR
AssertTrue(Condition := bOk, Message := 'all outputs finite at the zenith');
TEST_FINISHED();
END_METHOD

METHOD PRIVATE Zenith_Velocity_Is_Sidereal
VAR
	fbModel	: FB_PointingModelForward;
END_VAR
TEST('Zenith_Velocity_Is_Sidereal');
// at the site zenith the HA velocity is close to sidereal (0.0039 deg/s) and the Dec velocity is small, no jump (#4)
fbModel(HourAngle := 0.0, Declination := 51.5592378, Latitude := 51.5592378);
AssertEquals_LREAL(Expected := 0.003906120536459564, Actual := fbModel.HourAngle_velocity, Delta := 1.0E-9, Message := 'HA velocity');
AssertEquals_LREAL(Expected := 0.0000671134505799, Actual := fbModel.Declination_velocity, Delta := 1.0E-9, Message := 'Dec velocity');
TEST_FINISHED();
END_METHOD

METHOD PRIVATE Near_Zenith_Is_Continuous
VAR
	fbModel	: FB_PointingModelForward;
	fHaVelZenith	: LREAL;
	fDecVelZenith	: LREAL;
END_VAR
TEST('Near_Zenith_Is_Continuous');
fbModel(HourAngle := 0.0, Declination := 51.5592378, Latitude := 51.5592378);
fHaVelZenith := fbModel.HourAngle_velocity;
fDecVelZenith := fbModel.Declination_velocity;
fbModel(HourAngle := 1.0E-3, Declination := 51.5592378, Latitude := 51.5592378);
AssertEquals_LREAL(Expected := fHaVelZenith, Actual := fbModel.HourAngle_velocity, Delta := 1.0E-6, Message := 'HA velocity, HA offset');
AssertEquals_LREAL(Expected := fDecVelZenith, Actual := fbModel.Declination_velocity, Delta := 1.0E-6, Message := 'Dec velocity, HA offset');
fbModel(HourAngle := 0.0, Declination := 51.5592378 - 1.0E-3, Latitude := 51.5592378);
AssertEquals_LREAL(Expected := fHaVelZenith, Actual := fbModel.HourAngle_velocity, Delta := 1.0E-6, Message := 'HA velocity, Dec offset');
AssertEquals_LREAL(Expected := fDecVelZenith, Actual := fbModel.Declination_velocity, Delta := 1.0E-6, Message := 'Dec velocity, Dec offset');
TEST_FINISHED();
END_METHOD

METHOD PRIVATE Reference_Points_Unchanged
VAR
	fbModel	: FB_PointingModelForward;
END_VAR
TEST('Reference_Points_Unchanged');
// reference values from testing/check_pointing_zenith.py, site latitude
fbModel(HourAngle := 20.0, Declination := 40.0, Latitude := 51.5592378);
AssertEquals_LREAL(Expected := 0.2519851785590655, Actual := fbModel.HourAngle_correction, Delta := 1.0E-9, Message := 'HA correction 1');
AssertEquals_LREAL(Expected := -0.21403018480072264, Actual := fbModel.Declination_correction, Delta := 1.0E-9, Message := 'Dec correction 1');
AssertEquals_LREAL(Expected := 0.004006846115724003, Actual := fbModel.HourAngle_velocity, Delta := 1.0E-9, Message := 'HA velocity 1');
AssertEquals_LREAL(Expected := 0.00016906699168115099, Actual := fbModel.Declination_velocity, Delta := 1.0E-9, Message := 'Dec velocity 1');
fbModel(HourAngle := -35.0, Declination := 10.0, Latitude := 51.5592378);
AssertEquals_LREAL(Expected := 0.3090530046351645, Actual := fbModel.HourAngle_correction, Delta := 1.0E-9, Message := 'HA correction 2');
AssertEquals_LREAL(Expected := -0.19901388936334252, Actual := fbModel.Declination_correction, Delta := 1.0E-9, Message := 'Dec correction 2');
AssertEquals_LREAL(Expected := 0.00406630604072863, Actual := fbModel.HourAngle_velocity, Delta := 1.0E-9, Message := 'HA velocity 2');
AssertEquals_LREAL(Expected := -0.0001359293011053651, Actual := fbModel.Declination_velocity, Delta := 1.0E-9, Message := 'Dec velocity 2');
TEST_FINISHED();
END_METHOD

END_FUNCTION_BLOCK

// ---- POUs/FB_IagRig_Tests.TcPOU
// Spike S0 of the telescope state machine plan (BROTLib specs/plans/2026-10-21-telescope-state-machine-unification.md, step 0.3):
// can the real IAG50cm FB_TelescopeControl run on axis mocks that subclass FB_HourAngleControl/FB_DeclinationControl? The
// unlinked cabinet contacts read FALSE, which is a cabinet error and therefore a telescope error in every test: the rig sets
// them TRUE through pointers each scan (no production change).
FUNCTION_BLOCK FB_IagRig_Tests EXTENDS TcUnit.FB_TestSuite
VAR
	fbComm			: FB_NullComm;
	fbHa			: FB_HourAngleMock(comm := fbComm);
	fbDec			: FB_DeclinationMock(comm := fbComm);
	fbFocus			: FB_FocusMock;
	fbCovers		: FB_CoversMock;
	fbDome			: FB_DomeMock;
	fbTel			: FB_TelescopeControl(comm := fbComm);
	pBool			: POINTER TO BOOL;
END_VAR
VAR CONSTANT
	telescopeConfig	: ST_TelescopeConfig := (longitude := 9.9452433, latitude := 51.5592378, altitude := 100.0,
											 houranglePark := 0.0, declinationPark := 52.0, focusPark := 16.3,
											 hourangleHome := 0.0, declinationHome := 52.0, focusHome := 16.3,
											 name := 'Emmy Noether', diameter := 0.5, cabinet := 'Beckhoff', manufacturer := 'test',
											 mountOptions := 'HA-DEC', mount := 'HA_DEC');
END_VAR

Mock_Axis_Move_Reports_MoveDone();
Rig_Instantiates_Iag_Telescope();

METHOD PRIVATE CabinetOk
// the five contacts the cabinet error is made of (FB_CabinetControl, #10)
pBool := ADR(fbTel.fbCabinet.bAuxiliaryContact24V);		pBool^ := TRUE;
pBool := ADR(fbTel.fbCabinet.bAuxiliaryContact48V);		pBool^ := TRUE;
pBool := ADR(fbTel.fbCabinet.bAuxiliaryContactHADEC);	pBool^ := TRUE;
pBool := ADR(fbTel.fbCabinet.bAuxiliaryContactFOCUS);	pBool^ := TRUE;
pBool := ADR(fbTel.fbCabinet.bCollectiveReport24VFuse);	pBool^ := TRUE;
END_METHOD

METHOD PRIVATE Mock_Axis_Move_Reports_MoveDone
VAR
	i			: INT;
	bSeenDone	: BOOL;
END_VAR
TEST('Mock_Axis_Move_Reports_MoveDone');
fbHa.bEnable := TRUE;
FOR i := 1 TO 10 DO
	fbHa();
END_FOR
AssertTrue(Condition := fbHa.Ready, Message := 'enabled mock axis is ready');
AssertTrue(Condition := fbHa.Calibrated, Message := 'an enabled mock axis homes itself, like the real body');

fbHa.nMockMoveScans := 4;	// the default move takes 60 scans (long enough to interrupt it in the scenario suites)
fbHa.Position := 30.0;
fbHa.MoveAxis := TRUE;
FOR i := 1 TO 20 DO
	fbHa();
	IF fbHa.MoveDone THEN
		bSeenDone := TRUE;
	END_IF
END_FOR
AssertTrue(Condition := bSeenDone, Message := 'MoveDone was reported');
AssertFalse(Condition := fbHa.MoveAxis, Message := 'the move level is cleared on MoveDone');
AssertEquals_LREAL(Expected := 30.0, Actual := fbHa.ActualPosition, Delta := 0.001, Message := 'position is the target');
TEST_FINISHED();
END_METHOD

METHOD PRIVATE Rig_Instantiates_Iag_Telescope
VAR
	i	: INT;
END_VAR
TEST('Rig_Instantiates_Iag_Telescope');
FOR i := 1 TO 10 DO
	CabinetOk();
	fbTel(
		fbHourAngle := fbHa,
		fbDeclination := fbDec,
		fbFocus := fbFocus,
		fbDome := fbDome,
		fbCovers := fbCovers,
		telescopeConfig := telescopeConfig);
	fbHa();
	fbDec();
END_FOR
AssertFalse(Condition := fbTel.bError, Message := 'telescope on mock axes reports no error');
TEST_FINISHED();
END_METHOD

END_FUNCTION_BLOCK

// ---- POUs/FB_NullComm.TcPOU
// Minimal I_Comm stub for tests: every Publish/PublishLog call is a no-op that reports success,
// so FBs under test can call fbComm.Publish(...) freely without a real MQTT connection.
FUNCTION_BLOCK FB_NullComm IMPLEMENTS BROTLib.I_Comm
VAR
END_VAR

METHOD Publish : BOOL
VAR_INPUT
	domain			: STRING(255) := 'environment';
	location		: STRING(255) := 'roof';
	parameter		: STRING(255);
	value			: STRING(255);
END_VAR
VAR_OUTPUT
	published	: BOOL;
END_VAR
Publish := TRUE;
published := TRUE;
END_METHOD

METHOD PublishLREAL : BOOL
VAR_INPUT
	domain			: STRING(255) := 'environment';
	location		: STRING(255) := 'roof';
	parameter		: STRING(255);
	value			: LREAL;
END_VAR
VAR_OUTPUT
	published	: BOOL;
END_VAR
PublishLREAL := TRUE;
published := TRUE;
END_METHOD

METHOD PublishINT : BOOL
VAR_INPUT
	domain			: STRING(255) := 'environment';
	location		: STRING(255) := 'roof';
	parameter		: STRING(255);
	value			: LINT;
END_VAR
VAR_OUTPUT
	published	: BOOL;
END_VAR
PublishINT := TRUE;
published := TRUE;
END_METHOD

METHOD PublishBOOL : BOOL
VAR_INPUT
	domain			: STRING(255) := 'environment';
	location		: STRING(255) := 'roof';
	parameter		: STRING(255);
	value			: BOOL;
END_VAR
VAR_OUTPUT
	published	: BOOL;
END_VAR
PublishBOOL := TRUE;
published := TRUE;
END_METHOD

METHOD PublishString : BOOL
VAR_INPUT
	domain			: STRING(255) := 'environment';
	location		: STRING(255) := 'roof';
	parameter		: STRING(255);
	value			: STRING(255);
END_VAR
VAR_OUTPUT
	published	: BOOL;
END_VAR
PublishString := TRUE;
published := TRUE;
END_METHOD

METHOD PublishLog : BOOL
VAR_INPUT
	level		: STRING(255) := 'INFO';
	message		: STRING(255);
END_VAR
VAR_OUTPUT
	published	: BOOL;
END_VAR
PublishLog := TRUE;
published := TRUE;
END_METHOD

END_FUNCTION_BLOCK

// ---- POUs/FB_HourAngleMock.TcPOU
// Mock of FB_HourAngleControl for the telescope state machine tests (BROTLib plan 2026-10-21-telescope-state-machine-unification D1).
FUNCTION_BLOCK FB_HourAngleMock EXTENDS FB_HourAngleControl
VAR_INPUT
	nMockHomeScans	: UINT := 3;	// scans the calibration sweep (homing) takes (#197)
	nMockMoveScans	: UINT := 60;	// scans a move takes (the telescope sees Busy meanwhile)
	nMockStopScans	: UINT := 3;	// scans an MC_Stop takes until Done
	bMockNoStopDone	: BOOL;			// #120: the mock stop never reports Done (SetStopWithoutDone of the rig)
	nMockStartScans	: UINT;			// scans from the move command until the axis reports InMotion (0 = at once)
END_VAR
VAR_OUTPUT
	nStopEdges		: UINT;			// stop requests the telescope made (rising edges of StopAxis)
	nResetEdges		: UINT;			// resets the telescope sent to the axis (Reset())
END_VAR
VAR
	fbCore	: FB_AxisMockCore;
	pBool	: POINTER TO BOOL;
	pLreal	: POINTER TO LREAL;
	bInjected	: BOOL;
	nInjectedId	: UDINT;
END_VAR

// No SUPER^(): the real body (MC_* blocks, FB_LatchHome, AXIS_REF) does not run. The real property setters (MoveAxis ->
// fbAxis.MoveTo(), StopAxis -> fbAxis.Stop(), HomeAxis) stay, so the telescope sees the real command interface. The real body
// homes an enabled, uncalibrated axis by itself; the model does the same (bHome := bEnable). The model writes what the
// telescope reads: the base outputs and, through pointers (FB_Axis outputs are not writable from outside), the nested fbAxis outputs.
fbCore(bEnable := bEnable, bHome := bEnable, bMove := bMoveAxis, bStop := bStopAxis, fTarget := fPosition,
	nHomeScans := nMockHomeScans, nMoveScans := nMockMoveScans, nStopScans := nMockStopScans, nStartScans := nMockStartScans, bSuppressStopDone := bMockNoStopDone);

pBool := ADR(fbAxis.Ready);			pBool^ := fbCore.bReady;
pBool := ADR(fbAxis.Calibrated);	pBool^ := fbCore.bCalibrated;
pBool := ADR(fbAxis.HomeDone);		pBool^ := fbCore.bCalibrated;
pBool := ADR(fbAxis.HomeActive);	pBool^ := fbCore.bHoming;
pBool := ADR(fbAxis.Homing);		pBool^ := fbCore.bHoming;
pBool := ADR(fbAxis.InMotion);		pBool^ := fbCore.bInMotion;
pBool := ADR(fbAxis.StandStill);	pBool^ := fbCore.bStandStill;
pBool := ADR(fbAxis.MoveDone);		pBool^ := fbCore.bMoveDone;
pBool := ADR(fbAxis.Stopping);		pBool^ := fbCore.bStopping;
pBool := ADR(fbAxis.StopDone);		pBool^ := fbCore.bStopDone;
pBool := ADR(fbAxis.Busy);			pBool^ := fbCore.bInMotion OR fbCore.bHoming;
pLreal := ADR(fbAxis.ActualPosition);	pLreal^ := fbCore.fPosition;

bReady := fbCore.bReady AND fbCore.bStandStill;
nStopEdges := fbCore.nStopEdges;
bCalibrated := fbCore.bCalibrated;
fActualPosition := fbCore.fPosition;

// the real control body clears the level on MoveDone, and bStopAxis on StopDone
IF fbCore.bMoveDone THEN
	bMoveAxis := FALSE;
END_IF
IF fbCore.bStopDone THEN
	bStopAxis := FALSE;
END_IF
// a reset clears the injected error at once (ResetDone) and is counted
IF bReset THEN
	nResetEdges := nResetEdges + 1;
	bReset := FALSE;
	bInjected := FALSE;
	nInjectedId := 0;
END_IF
bError := bInjected;
nErrorID := nInjectedId;

// the axis reports an error with this id until the telescope resets it (bError/nErrorID are what the telescope reads)
METHOD InjectError
VAR_INPUT
	nId	: UDINT;
END_VAR
bInjected := TRUE;
nInjectedId := nId;
END_METHOD

END_FUNCTION_BLOCK

// ---- POUs/FB_AxisMockCore.TcPOU
// Motion model of one mocked axis (telescope state machine mock rig, BROTLib plan 2026-10-21-telescope-state-machine-unification).
// One call = one PLC scan of the axis part. Enable -> Ready after nReadyScans, homing -> calibrated after nHomeScans, a rising
// bMove -> InMotion for nMoveScans, then MoveDone for one scan and the position is the target. Only the levels the telescope
// writes are inputs; nothing here touches an MC_* block. Same model as MONETcommonTests.
FUNCTION_BLOCK FB_AxisMockCore
VAR_INPUT
	bEnable			: BOOL;
	bHome			: BOOL;
	bMove			: BOOL;
	bStop			: BOOL;		// the StopAxis level: a rising edge is a stop request (MC_Stop)
	fTarget			: LREAL;
	nReadyScans		: UINT := 2;
	nHomeScans		: UINT := 3;
	nMoveScans		: UINT := 4;
	nStopScans		: UINT := 3;
	bSuppressStopDone	: BOOL;	// the stop ends at rest but bStopDone is never reported (a lost Done, #120)
	nStartScans		: UINT;		// scans between the move command and the axis reporting InMotion (the NC takes a few cycles; 0 = at once). #92
END_VAR
VAR_OUTPUT
	bReady			: BOOL;
	bCalibrated		: BOOL;
	bHoming			: BOOL;
	bInMotion		: BOOL;
	bStandStill		: BOOL := TRUE;
	bMoveDone		: BOOL;		// one scan
	bStopping		: BOOL;
	bStopDone		: BOOL;		// one scan
	nStopEdges		: UINT;		// rising edges of bStop, i.e. MC_Stop requests
	fPosition		: LREAL;
END_VAR
VAR
	nReadyCount		: UINT;
	nHomeCount		: UINT;
	nMoveCount		: UINT;
	nStopCount		: UINT;
	nStartCount		: UINT;
	bStartPending	: BOOL;
	rtMove			: R_TRIG;
	rtStop			: R_TRIG;
END_VAR

bMoveDone := FALSE;
bStopDone := FALSE;

// a stop request aborts a running move where it is (the model has no interpolation: the position stays) and takes
// nStopScans scans, then reports Done for one scan
rtStop(CLK := bStop);
IF rtStop.Q THEN
	nStopEdges := nStopEdges + 1;
	bStopping := TRUE;
	nStopCount := 0;
	bInMotion := FALSE;
	bStartPending := FALSE;
END_IF
IF bStopping THEN
	nStopCount := nStopCount + 1;
	IF nStopCount >= nStopScans THEN
		bStopping := FALSE;
		bStopDone := NOT bSuppressStopDone;
	END_IF
END_IF

IF bEnable THEN
	IF nReadyCount >= nReadyScans THEN
		bReady := TRUE;
	ELSE
		nReadyCount := nReadyCount + 1;
	END_IF
ELSE
	nReadyCount := 0;
	bReady := FALSE;
END_IF

IF bHome AND bReady AND NOT bCalibrated THEN
	bHoming := TRUE;
	nHomeCount := nHomeCount + 1;
	IF nHomeCount >= nHomeScans THEN
		bCalibrated := TRUE;
		bHoming := FALSE;
		nHomeCount := 0;
	END_IF
ELSE
	bHoming := FALSE;
END_IF

rtMove(CLK := bMove);
IF rtMove.Q AND bReady AND bCalibrated AND NOT bStopping THEN
	IF nStartScans = 0 THEN
		bInMotion := TRUE;
		nMoveCount := 0;
	ELSE
		// the move command is out, the axis still reports StandStill until the NC has started it (#92)
		bStartPending := TRUE;
		nStartCount := 0;
	END_IF
ELSIF bStartPending THEN
	nStartCount := nStartCount + 1;
	IF nStartCount >= nStartScans THEN
		bStartPending := FALSE;
		bInMotion := TRUE;
		nMoveCount := 0;
	END_IF
END_IF
IF bInMotion THEN
	nMoveCount := nMoveCount + 1;
	IF nMoveCount >= nMoveScans THEN
		fPosition := fTarget;
		bInMotion := FALSE;
		bMoveDone := TRUE;
	END_IF
END_IF

bStandStill := NOT bInMotion AND NOT bHoming AND NOT bStopping;

END_FUNCTION_BLOCK

// ---- POUs/FB_DeclinationMock.TcPOU
// Mock of FB_DeclinationControl for the telescope state machine tests (BROTLib plan 2026-10-21-telescope-state-machine-unification D1).
FUNCTION_BLOCK FB_DeclinationMock EXTENDS FB_DeclinationControl
VAR_INPUT
	nMockHomeScans	: UINT := 3;	// scans the calibration sweep (homing) takes (#197)
	nMockMoveScans	: UINT := 60;	// scans a move takes (the telescope sees Busy meanwhile)
	nMockStopScans	: UINT := 3;	// scans an MC_Stop takes until Done
	bMockNoStopDone	: BOOL;			// #120: the mock stop never reports Done (SetStopWithoutDone of the rig)
	nMockStartScans	: UINT;			// scans from the move command until the axis reports InMotion (0 = at once)
END_VAR
VAR_OUTPUT
	nStopEdges		: UINT;			// stop requests the telescope made (rising edges of StopAxis)
	nResetEdges		: UINT;			// resets the telescope sent to the axis (Reset())
END_VAR
VAR
	fbCore	: FB_AxisMockCore;
	pBool	: POINTER TO BOOL;
	pLreal	: POINTER TO LREAL;
	bInjected	: BOOL;
	nInjectedId	: UDINT;
END_VAR

// No SUPER^(): the real body (MC_* blocks, FB_LatchHome, AXIS_REF) does not run. The real property setters (MoveAxis ->
// fbAxis.MoveTo(), StopAxis -> fbAxis.Stop(), HomeAxis) stay, so the telescope sees the real command interface. The real body
// homes an enabled, uncalibrated axis by itself; the model does the same (bHome := bEnable). The model writes what the
// telescope reads: the base outputs and, through pointers (FB_Axis outputs are not writable from outside), the nested fbAxis outputs.
fbCore(bEnable := bEnable, bHome := bEnable, bMove := bMoveAxis, bStop := bStopAxis, fTarget := fPosition,
	nHomeScans := nMockHomeScans, nMoveScans := nMockMoveScans, nStopScans := nMockStopScans, nStartScans := nMockStartScans, bSuppressStopDone := bMockNoStopDone);

pBool := ADR(fbAxis.Ready);			pBool^ := fbCore.bReady;
pBool := ADR(fbAxis.Calibrated);	pBool^ := fbCore.bCalibrated;
pBool := ADR(fbAxis.HomeDone);		pBool^ := fbCore.bCalibrated;
pBool := ADR(fbAxis.HomeActive);	pBool^ := fbCore.bHoming;
pBool := ADR(fbAxis.Homing);		pBool^ := fbCore.bHoming;
pBool := ADR(fbAxis.InMotion);		pBool^ := fbCore.bInMotion;
pBool := ADR(fbAxis.StandStill);	pBool^ := fbCore.bStandStill;
pBool := ADR(fbAxis.MoveDone);		pBool^ := fbCore.bMoveDone;
pBool := ADR(fbAxis.Stopping);		pBool^ := fbCore.bStopping;
pBool := ADR(fbAxis.StopDone);		pBool^ := fbCore.bStopDone;
pBool := ADR(fbAxis.Busy);			pBool^ := fbCore.bInMotion OR fbCore.bHoming;
pLreal := ADR(fbAxis.ActualPosition);	pLreal^ := fbCore.fPosition;

bReady := fbCore.bReady AND fbCore.bStandStill;
nStopEdges := fbCore.nStopEdges;
bCalibrated := fbCore.bCalibrated;
fActualPosition := fbCore.fPosition;

// the real control body clears the level on MoveDone, and bStopAxis on StopDone
IF fbCore.bMoveDone THEN
	bMoveAxis := FALSE;
END_IF
IF fbCore.bStopDone THEN
	bStopAxis := FALSE;
END_IF
// a reset clears the injected error at once (ResetDone) and is counted
IF bReset THEN
	nResetEdges := nResetEdges + 1;
	bReset := FALSE;
	bInjected := FALSE;
	nInjectedId := 0;
END_IF
bError := bInjected;
nErrorID := nInjectedId;

// the axis reports an error with this id until the telescope resets it (bError/nErrorID are what the telescope reads)
METHOD InjectError
VAR_INPUT
	nId	: UDINT;
END_VAR
bInjected := TRUE;
nInjectedId := nId;
END_METHOD

END_FUNCTION_BLOCK

// ---- POUs/FB_FocusMock.TcPOU
// Mock of the focus axis (I_Focus) for the telescope state machine tests: enabled = ready and calibrated at once (the telescope never sets HomeAxis), the
// position follows the target at once. Status only, no motion model.
FUNCTION_BLOCK FB_FocusMock IMPLEMENTS BROTLib.I_Focus
VAR
	bEn		: BOOL;
	bCal	: BOOL;
	bHome	: BOOL;
	bNeg	: BOOL;
	bPos	: BOOL;
	fPos	: LREAL;
	fTarget	: LREAL;
	fVel	: LREAL;
	nStop	: INT;		// number of Stop() calls
END_VAR

IF bEn THEN
	bCal := TRUE;
END_IF
fPos := fTarget;

METHOD Stop : BOOL
nStop := nStop + 1;
Stop := TRUE;
END_METHOD

PROPERTY MinPosition : LREAL
GET
MinPosition := -1.0E6;
END_GET
END_PROPERTY

PROPERTY MaxPosition : LREAL
GET
MaxPosition := 1.0E6;
END_GET
END_PROPERTY

METHOD Reset : BOOL
Reset := TRUE;
END_METHOD

PROPERTY ActualPosition : LREAL
GET
ActualPosition := fPos;
END_GET
SET
fPos := ActualPosition;
END_SET
END_PROPERTY

PROPERTY Busy : BOOL
GET
Busy := FALSE;
END_GET
END_PROPERTY

PROPERTY Calibrated : BOOL
GET
Calibrated := bCal;
END_GET
END_PROPERTY

PROPERTY Enable : BOOL
GET
Enable := bEn;
END_GET
SET
bEn := Enable;
END_SET
END_PROPERTY

PROPERTY Error : BOOL
GET
Error := FALSE;
END_GET
END_PROPERTY

PROPERTY ErrorID : UDINT
GET
ErrorID := 0;
END_GET
END_PROPERTY

PROPERTY HomeAxis : BOOL
GET
HomeAxis := bHome;
END_GET
SET
bHome := HomeAxis;
END_SET
END_PROPERTY

PROPERTY InNegLimit : BOOL
GET
InNegLimit := FALSE;
END_GET
END_PROPERTY

PROPERTY InPosLimit : BOOL
GET
InPosLimit := FALSE;
END_GET
END_PROPERTY

PROPERTY MoveNeg : BOOL
GET
MoveNeg := bNeg;
END_GET
SET
bNeg := MoveNeg;
END_SET
END_PROPERTY

PROPERTY MovePos : BOOL
GET
MovePos := bPos;
END_GET
SET
bPos := MovePos;
END_SET
END_PROPERTY

PROPERTY Position : LREAL
GET
Position := fTarget;
END_GET
SET
fTarget := Position;
END_SET
END_PROPERTY

PROPERTY Ready : BOOL
GET
Ready := bEn;
END_GET
END_PROPERTY

PROPERTY Velocity : LREAL
GET
Velocity := fVel;
END_GET
SET
fVel := Velocity;
END_SET
END_PROPERTY

END_FUNCTION_BLOCK

// ---- POUs/FB_CoversMock.TcPOU
// Mock of the mirror covers (I_MirrorCovers): Open/Close take effect at once, unless bHoldClose is set: then Close is only counted
// and the covers stay open until the test sets bClosed (a slow closing, IAG50cm#187).
FUNCTION_BLOCK FB_CoversMock IMPLEMENTS BROTLib.I_MirrorCovers
VAR
	bOpened		: BOOL;
	bClosed		: BOOL := TRUE;
	bFailed		: BOOL;
	bHoldClose	: BOOL;
	nOpenCalls	: UINT;
	nCloseCalls	: UINT;
END_VAR

METHOD Open : BOOL
bOpened := TRUE;
bClosed := FALSE;
nOpenCalls := nOpenCalls + 1;
Open := TRUE;
END_METHOD

METHOD Close : BOOL
bOpened := FALSE;
IF NOT bHoldClose THEN
	bClosed := TRUE;
END_IF
nCloseCalls := nCloseCalls + 1;
Close := TRUE;
END_METHOD

// while bHold is TRUE a Close() is only counted and the covers stay open (a slow closing, IAG50cm#187)
METHOD HoldClose
VAR_INPUT
	bHold	: BOOL;
END_VAR
bHoldClose := bHold;
END_METHOD

// the held closing is done: the covers are closed now
METHOD FinishClose
bHoldClose := FALSE;
bOpened := FALSE;
bClosed := TRUE;
END_METHOD

METHOD Reset : BOOL
bFailed := FALSE;
Reset := TRUE;
END_METHOD

PROPERTY Opened : BOOL
GET
Opened := bOpened;
END_GET
END_PROPERTY

PROPERTY Closed : BOOL
GET
Closed := bClosed;
END_GET
END_PROPERTY

PROPERTY Error : BOOL
GET
Error := bFailed;
END_GET
END_PROPERTY

END_FUNCTION_BLOCK

// ---- POUs/FB_DomeMock.TcPOU
// Mock of the dome (I_Dome): the commands only count, nothing moves.
FUNCTION_BLOCK FB_DomeMock IMPLEMENTS BROTLib.I_Dome
VAR
	bFailed		: BOOL;
	bIsParked	: BOOL := TRUE;
	bIsTracking	: BOOL;
	fPos		: LREAL;
	eShutter	: BROTLib.E_RoofState;
	nParkCalls	: UINT;
	nTrackCalls	: UINT;
END_VAR

METHOD Close : BOOL
Close := TRUE;
END_METHOD

METHOD Open : BOOL
Open := TRUE;
END_METHOD

METHOD Park : BOOL
nParkCalls := nParkCalls + 1;
bIsParked := TRUE;
bIsTracking := FALSE;
Park := TRUE;
END_METHOD

METHOD Reset : BOOL
bFailed := FALSE;
Reset := TRUE;
END_METHOD

METHOD Stop : BOOL
Stop := TRUE;
END_METHOD

METHOD StopTrack : BOOL
bIsTracking := FALSE;
StopTrack := TRUE;
END_METHOD

METHOD Track : BOOL
nTrackCalls := nTrackCalls + 1;
bIsParked := FALSE;
bIsTracking := TRUE;
Track := TRUE;
END_METHOD

PROPERTY Capabilities : INT
GET
Capabilities := 0;
END_GET
END_PROPERTY

PROPERTY Error : BOOL
GET
Error := bFailed;
END_GET
END_PROPERTY

PROPERTY ErrorID : UDINT
GET
ErrorID := 0;
END_GET
END_PROPERTY

PROPERTY Parked : BOOL
GET
Parked := bIsParked;
END_GET
END_PROPERTY

PROPERTY Position : LREAL
GET
Position := fPos;
END_GET
SET
fPos := Position;
END_SET
END_PROPERTY

PROPERTY RotState : BROTLib.E_DomeRotationState
GET
RotState := BROTLib.E_DomeRotationState.idle;
END_GET
END_PROPERTY

PROPERTY ShutterState : BROTLib.E_RoofState
GET
ShutterState := eShutter;
END_GET
SET
eShutter := ShutterState;
END_SET
END_PROPERTY

PROPERTY Tracking : BOOL
GET
Tracking := bIsTracking;
END_GET
END_PROPERTY

END_FUNCTION_BLOCK

// ---- POUs/IagStopDuringSlew_Tests.TcPOU
// Characterization of FB_TelescopeControl (IAG50cm) for a stop during a slew, on mock axes (plan step 2, IAG50cmTests README).
// These tests pin what the code does today, with the line of the behaviour in a comment; they are not a specification. Every
// test owns a rig and runs over many PLC cycles (VAR_INST of the method, one Scan() per cycle); TcUnit calls all test methods
// every cycle, so the rigs warm up their clocks in parallel. A step that does not happen within its cycle budget fails the
// test with a message instead of hanging the run.
FUNCTION_BLOCK IagStopDuringSlew_Tests EXTENDS TcUnit.FB_TestSuite
VAR
END_VAR

Stop_During_Slew_One_Stop_For_The_Moving_Axis();
Stop_Drops_The_Move_Before_Sending_The_Axis_Stop();
Stop_Clears_The_Slew_And_Settles();

// #108: one MC_Stop per axis that is not at rest, none for an axis at rest. The IAG slew moves one axis at a time
// (_SlewTelescope stages 30..33 / 40..43), so only one axis is moving when the stop comes.
METHOD PRIVATE Stop_During_Slew_One_Stop_For_The_Moving_Axis
VAR_INST
	rig			: FB_IagRig;
	nStep		: INT;
	nCycles		: UINT;
	bHaMoving	: BOOL;
	sTest		: STRING(80);
END_VAR
TEST('Stop_During_Slew_One_Stop_For_The_Moving_Axis');
sTest := 'Stop_During_Slew_One_Stop_For_The_Moving_Axis: ';
IF nStep >= 90 THEN
	RETURN;
END_IF
rig.Scan();
nCycles := nCycles + 1;
CASE nStep OF
0:	// wait for the clock, then power on
	IF rig.ClockValid THEN
		rig.fbTel.Init();
		nStep := 10;
		nCycles := 0;
	ELSIF nCycles > 2000 THEN
		AssertTrue(Condition := FALSE, Message := 'the astronomical clock never became valid');
		F_Note(bFailed := NOT (FALSE), sText := CONCAT(sTest, 'the astronomical clock never became valid'));
		nStep := 99;
		TEST_FINISHED();
	END_IF
10:	// wait until the startup has finished (READY_STATE 1.0), then slew
	IF rig.Online THEN
		rig.fbTel.Slew(fAzimuth := 180.0, fAltitude := 45.0);
		nStep := 20;
		nCycles := 0;
	ELSIF nCycles > 1500 THEN
		AssertTrue(Condition := FALSE, Message := 'the mock telescope did not reach READY_STATE 1.0');
		F_Note(bFailed := NOT (FALSE), sText := CONCAT(sTest, 'the mock telescope did not reach READY_STATE 1.0'));
		nStep := 99;
		TEST_FINISHED();
	END_IF
20:	// wait until one axis is moving (the slew moves HA and Dec one after the other)
	IF rig.fbHa.MoveAxis OR rig.fbDec.MoveAxis THEN
		bHaMoving := rig.fbHa.MoveAxis;
		AssertTrue(Condition := rig.fbTel.bSlewActive, Message := 'bSlew is set while the slew runs');
		F_Note(bFailed := NOT (rig.fbTel.bSlewActive), sText := CONCAT(sTest, 'bSlew is set while the slew runs'));
		// IAG50cm#17 step 0.3: the coordinate chain runs inside the telescope (the migration must keep it running). The slew
		// target az 180 / alt 45 is on the meridian: Dec about latitude - 45 = 6.56 deg, hour angle about 0.
		AssertFalse(Condition := F_NoteNear(CONCAT(sTest, 'Julian date'), 2461000.0, rig.fbTel.fJd, 2000.0), Message := 'fJd follows the clock');
		AssertFalse(Condition := F_NoteNear(CONCAT(sTest, 'slew target Dec'), 51.5592378 - 45.0, rig.fbTel.fDeclinationCalc, 0.5), Message := 'slew target declination');
		AssertTrue(Condition := COS(rig.fbTel.fHourAngleCalc * 0.017453292519943295) > 0.9999, Message := 'slew target hour angle about 0');
		F_Note(bFailed := NOT (COS(rig.fbTel.fHourAngleCalc * 0.017453292519943295) > 0.9999), sText := CONCAT(sTest, 'slew target hour angle about 0'));
		AssertTrue(Condition := ABS(rig.fbTel.fDeclinationApparent) <= 90.0, Message := 'apparent declination is finite');
		F_Note(bFailed := NOT (ABS(rig.fbTel.fDeclinationApparent) <= 90.0), sText := CONCAT(sTest, 'apparent declination is finite'));
		AssertTrue(Condition := ABS(rig.fbTel.fElevationCalc) <= 90.0, Message := 'target elevation is finite');
		F_Note(bFailed := NOT (ABS(rig.fbTel.fElevationCalc) <= 90.0), sText := CONCAT(sTest, 'target elevation is finite'));
		nStep := 30;
		nCycles := 0;
	ELSIF nCycles > 300 THEN
		AssertTrue(Condition := FALSE, Message := 'the slew did not start an axis move');
		F_Note(bFailed := NOT (FALSE), sText := CONCAT(sTest, 'the slew did not start an axis move'));
		nStep := 99;
		TEST_FINISHED();
	END_IF
30:	// let the move run for a few scans, then stop
	IF nCycles >= 5 THEN
		rig.fbTel.Stop();
		nStep := 40;
		nCycles := 0;
	END_IF
40:	// wait until the stop has settled
	IF NOT rig.fbTel.bStopActive AND rig.fbTel.bStopped AND nCycles > 5 THEN
		AssertEquals_UINT(Expected := SEL(bHaMoving, UINT#0, UINT#1), Actual := rig.fbHa.nStopEdges, Message := 'HA: one stop if it was the moving axis, none otherwise');
		F_Note(bFailed := (SEL(bHaMoving, UINT#0, UINT#1)) <> (rig.fbHa.nStopEdges), sText := CONCAT(sTest, 'HA: one stop if it was the moving axis, none otherwise'));
		AssertEquals_UINT(Expected := SEL(bHaMoving, UINT#1, UINT#0), Actual := rig.fbDec.nStopEdges, Message := 'Dec: one stop if it was the moving axis, none otherwise');
		F_Note(bFailed := (SEL(bHaMoving, UINT#1, UINT#0)) <> (rig.fbDec.nStopEdges), sText := CONCAT(sTest, 'Dec: one stop if it was the moving axis, none otherwise'));
		nStep := 99;
		TEST_FINISHED();
	ELSIF nCycles > 400 THEN
		AssertTrue(Condition := FALSE, Message := 'the stop did not settle');
		F_Note(bFailed := NOT (FALSE), sText := CONCAT(sTest, 'the stop did not settle'));
		nStep := 99;
		TEST_FINISHED();
	END_IF
END_CASE
END_METHOD

// _StopTelescope (I:1927-1953): the first scan of a stop only drops MoveAxis (the first branch; that does not stop a running
// move); the axis stop (StopAxis) is sent in the next scan.
METHOD PRIVATE Stop_Drops_The_Move_Before_Sending_The_Axis_Stop
VAR_INST
	rig			: FB_IagRig;
	nStep		: INT;
	nCycles		: UINT;
	bHaMoving	: BOOL;
	sTest		: STRING(80);
END_VAR
TEST('Stop_Drops_The_Move_Before_Sending_The_Axis_Stop');
sTest := 'Stop_Drops_The_Move_Before_Sending_The_Axis_Stop: ';
IF nStep >= 90 THEN
	RETURN;
END_IF
rig.Scan();
nCycles := nCycles + 1;
CASE nStep OF
0:	// wait for the clock, then power on
	IF rig.ClockValid THEN
		rig.fbTel.Init();
		nStep := 10;
		nCycles := 0;
	ELSIF nCycles > 2000 THEN
		AssertTrue(Condition := FALSE, Message := 'the astronomical clock never became valid');
		F_Note(bFailed := NOT (FALSE), sText := CONCAT(sTest, 'the astronomical clock never became valid'));
		nStep := 99;
		TEST_FINISHED();
	END_IF
10:	// wait until the startup has finished (READY_STATE 1.0), then slew
	IF rig.Online THEN
		rig.fbTel.Slew(fAzimuth := 180.0, fAltitude := 45.0);
		nStep := 20;
		nCycles := 0;
	ELSIF nCycles > 1500 THEN
		AssertTrue(Condition := FALSE, Message := 'the mock telescope did not reach READY_STATE 1.0');
		F_Note(bFailed := NOT (FALSE), sText := CONCAT(sTest, 'the mock telescope did not reach READY_STATE 1.0'));
		nStep := 99;
		TEST_FINISHED();
	END_IF
20:	// wait until one axis is moving (the slew moves HA and Dec one after the other)
	IF rig.fbHa.MoveAxis OR rig.fbDec.MoveAxis THEN
		bHaMoving := rig.fbHa.MoveAxis;
		AssertTrue(Condition := rig.fbTel.bSlewActive, Message := 'bSlew is set while the slew runs');
		F_Note(bFailed := NOT (rig.fbTel.bSlewActive), sText := CONCAT(sTest, 'bSlew is set while the slew runs'));
		nStep := 30;
		nCycles := 0;
	ELSIF nCycles > 300 THEN
		AssertTrue(Condition := FALSE, Message := 'the slew did not start an axis move');
		F_Note(bFailed := NOT (FALSE), sText := CONCAT(sTest, 'the slew did not start an axis move'));
		nStep := 99;
		TEST_FINISHED();
	END_IF
30:	// let the move run for a few scans, then stop
	IF nCycles >= 5 THEN
		rig.fbTel.Stop();
		nStep := 40;
		nCycles := 0;
	END_IF
40:	// scan 1 of the stop has just run: the move is dropped, no axis stop yet; scan 2 sends it
	IF nCycles = 1 THEN
		AssertFalse(Condition := rig.fbHa.MoveAxis OR rig.fbDec.MoveAxis, Message := 'scan 1 of the stop drops the move');
		F_Note(bFailed := (rig.fbHa.MoveAxis OR rig.fbDec.MoveAxis), sText := CONCAT(sTest, 'scan 1 of the stop drops the move'));
		AssertFalse(Condition := rig.fbHa.StopAxis OR rig.fbDec.StopAxis, Message := 'scan 1 of the stop does not send an axis stop yet');
		F_Note(bFailed := (rig.fbHa.StopAxis OR rig.fbDec.StopAxis), sText := CONCAT(sTest, 'scan 1 of the stop does not send an axis stop yet'));
	ELSIF nCycles = 2 THEN
		AssertTrue(Condition := SEL(bHaMoving, rig.fbDec.StopAxis, rig.fbHa.StopAxis), Message := 'scan 2 sends the stop to the axis that was moving');
		F_Note(bFailed := NOT (SEL(bHaMoving, rig.fbDec.StopAxis, rig.fbHa.StopAxis)), sText := CONCAT(sTest, 'scan 2 sends the stop to the axis that was moving'));
		AssertFalse(Condition := SEL(bHaMoving, rig.fbHa.StopAxis, rig.fbDec.StopAxis), Message := 'scan 2 sends no stop to the axis at rest');
		F_Note(bFailed := (SEL(bHaMoving, rig.fbHa.StopAxis, rig.fbDec.StopAxis)), sText := CONCAT(sTest, 'scan 2 sends no stop to the axis at rest'));
		nStep := 99;
		TEST_FINISHED();
	END_IF
END_CASE
END_METHOD

// Arbitration (I:501-526): a user stop during a slew drops bSlew, runs the stop until the axes stand still, and releases bStop.
METHOD PRIVATE Stop_Clears_The_Slew_And_Settles
VAR_INST
	rig			: FB_IagRig;
	nStep		: INT;
	nCycles		: UINT;
	bHaMoving	: BOOL;
	sTest		: STRING(80);
END_VAR
TEST('Stop_Clears_The_Slew_And_Settles');
sTest := 'Stop_Clears_The_Slew_And_Settles: ';
IF nStep >= 90 THEN
	RETURN;
END_IF
rig.Scan();
nCycles := nCycles + 1;
CASE nStep OF
0:	// wait for the clock, then power on
	IF rig.ClockValid THEN
		rig.fbTel.Init();
		nStep := 10;
		nCycles := 0;
	ELSIF nCycles > 2000 THEN
		AssertTrue(Condition := FALSE, Message := 'the astronomical clock never became valid');
		F_Note(bFailed := NOT (FALSE), sText := CONCAT(sTest, 'the astronomical clock never became valid'));
		nStep := 99;
		TEST_FINISHED();
	END_IF
10:	// wait until the startup has finished (READY_STATE 1.0), then slew
	IF rig.Online THEN
		rig.fbTel.Slew(fAzimuth := 180.0, fAltitude := 45.0);
		nStep := 20;
		nCycles := 0;
	ELSIF nCycles > 1500 THEN
		AssertTrue(Condition := FALSE, Message := 'the mock telescope did not reach READY_STATE 1.0');
		F_Note(bFailed := NOT (FALSE), sText := CONCAT(sTest, 'the mock telescope did not reach READY_STATE 1.0'));
		nStep := 99;
		TEST_FINISHED();
	END_IF
20:	// wait until one axis is moving (the slew moves HA and Dec one after the other)
	IF rig.fbHa.MoveAxis OR rig.fbDec.MoveAxis THEN
		bHaMoving := rig.fbHa.MoveAxis;
		AssertTrue(Condition := rig.fbTel.bSlewActive, Message := 'bSlew is set while the slew runs');
		F_Note(bFailed := NOT (rig.fbTel.bSlewActive), sText := CONCAT(sTest, 'bSlew is set while the slew runs'));
		nStep := 30;
		nCycles := 0;
	ELSIF nCycles > 300 THEN
		AssertTrue(Condition := FALSE, Message := 'the slew did not start an axis move');
		F_Note(bFailed := NOT (FALSE), sText := CONCAT(sTest, 'the slew did not start an axis move'));
		nStep := 99;
		TEST_FINISHED();
	END_IF
30:	// let the move run for a few scans, then stop
	IF nCycles >= 5 THEN
		rig.fbTel.Stop();
		nStep := 40;
		nCycles := 0;
	END_IF
40:
	IF NOT rig.fbTel.bStopActive AND rig.fbTel.bStopped AND nCycles > 5 THEN
		AssertFalse(Condition := rig.fbTel.bSlewActive, Message := 'the stop dropped bSlew');
		F_Note(bFailed := (rig.fbTel.bSlewActive), sText := CONCAT(sTest, 'the stop dropped bSlew'));
		AssertFalse(Condition := rig.fbHa.MoveAxis OR rig.fbDec.MoveAxis, Message := 'no axis move is left');
		F_Note(bFailed := (rig.fbHa.MoveAxis OR rig.fbDec.MoveAxis), sText := CONCAT(sTest, 'no axis move is left'));
		AssertTrue(Condition := rig.fbTel.bReady, Message := 'the telescope is still ready after the stop');
		F_Note(bFailed := NOT (rig.fbTel.bReady), sText := CONCAT(sTest, 'the telescope is still ready after the stop'));
		nStep := 99;
		TEST_FINISHED();
	ELSIF nCycles > 400 THEN
		AssertTrue(Condition := FALSE, Message := 'the stop did not settle');
		F_Note(bFailed := NOT (FALSE), sText := CONCAT(sTest, 'the stop did not settle'));
		nStep := 99;
		TEST_FINISHED();
	END_IF
END_CASE
END_METHOD

END_FUNCTION_BLOCK

// ---- POUs/FB_IagRig.TcPOU
// The IAG50cm telescope on mock axes, scanned in the MAIN order (axes, then the telescope; IAG50cm/POUs/MAIN.TcPOU).
// One Scan() is one PLC scan. The scenario tests own one rig each (VAR_INST of the test method) and call Scan() once per
// PLC cycle: the astronomical clock needs a real NT_GetTime round trip (up to about 5 s) before FB_TelescopeControl accepts a
// goto/slew/track, so a rig is not usable before ClockValid. Everything else counts scans, not time.
// Plan: BROTLib specs/plans/2026-10-21-telescope-state-machine-unification.md (D1, step 2).
FUNCTION_BLOCK FB_IagRig
VAR
	fbComm			: FB_RecordingComm;	// records nothing until a test calls Start (IagTelemetry_Tests)
	fbHa			: FB_HourAngleMock(comm := fbComm);
	fbDec			: FB_DeclinationMock(comm := fbComm);
	fbFocus			: FB_FocusMock;
	fbCovers		: FB_CoversMock;
	fbDome			: FB_DomeMock;
	fbTel			: FB_TelescopeControl(comm := fbComm);
	pBool			: POINTER TO BOOL;
	nScans			: UDINT;
	nTimeDivisor	: UDINT := 1;	// the time seam of the telescope under test (SetTimeDivisor)
	fHorizon		: LREAL := 1.0;	// the horizon limit passed to the telescope (an input, so tests set it here; #84)
END_VAR
VAR CONSTANT
	telescopeConfig	: ST_TelescopeConfig := (longitude := 9.9452433, latitude := 51.5592378, altitude := 100.0,
											 houranglePark := 0.0, declinationPark := 52.0, focusPark := 16.3,
											 hourangleHome := 0.0, declinationHome := 52.0, focusHome := 16.3,
											 name := 'Emmy Noether', diameter := 0.5, cabinet := 'Beckhoff', manufacturer := 'test',
											 mountOptions := 'HA-DEC', mount := 'HA_DEC');
END_VAR

METHOD Scan
// the five contacts the cabinet error is made of (FB_CabinetControl, #10); unlinked they read FALSE
pBool := ADR(fbTel.fbCabinet.bAuxiliaryContact24V);		pBool^ := TRUE;
pBool := ADR(fbTel.fbCabinet.bAuxiliaryContact48V);		pBool^ := TRUE;
pBool := ADR(fbTel.fbCabinet.bAuxiliaryContactHADEC);	pBool^ := TRUE;
pBool := ADR(fbTel.fbCabinet.bAuxiliaryContactFOCUS);	pBool^ := TRUE;
pBool := ADR(fbTel.fbCabinet.bCollectiveReport24VFuse);	pBool^ := TRUE;

fbHa();
fbDec();
fbFocus();
fbTel(
	fbHourAngle := fbHa,
	fbDeclination := fbDec,
	fbFocus := fbFocus,
	fbDome := fbDome,
	fbCovers := fbCovers,
	telescopeConfig := telescopeConfig,
	nTimeDivisor := nTimeDivisor,
	fHorizon := fHorizon);
nScans := nScans + 1;
END_METHOD

PROPERTY ClockValid : BOOL
GET
ClockValid := fbTel.fbTime.bValid;
END_GET
END_PROPERTY

PROPERTY Online : BOOL
GET
Online := fbTel.ReadyState = 1.0;
END_GET
END_PROPERTY

// divides every long timeout of the telescope (600 s, 2 min, 12 h) by nValue, for this rig only (1 = real times)
METHOD SetTimeDivisor
VAR_INPUT
	nValue	: UDINT;
END_VAR
nTimeDivisor := nValue;
fbTel.nTimeDivisor := nValue;
END_METHOD

// the horizon limit of the telescope under test (an input of the telescope, so it cannot be written from outside; #84)
METHOD SetHorizon
VAR_INPUT
	fValue	: LREAL;
END_VAR
fHorizon := fValue;
END_METHOD

// scans a move takes on both mock axes (default 60)
METHOD SetMoveScans
VAR_INPUT
	nScans	: UINT;
END_VAR
fbHa.nMockMoveScans := nScans;
fbDec.nMockMoveScans := nScans;
END_METHOD

// scans the calibration sweep (homing) of each mock axis takes (default 3, #197)
METHOD SetHomeScans
VAR_INPUT
	nHa		: UINT;
	nDec	: UINT;
END_VAR
fbHa.nMockHomeScans := nHa;
fbDec.nMockHomeScans := nDec;
END_METHOD

// scans from a move command until the mock axes report InMotion (default 0: at once); the NC on the real axes takes a few cycles
METHOD SetStartScans
VAR_INPUT
	nScans	: UINT;
END_VAR
fbHa.nMockStartScans := nScans;
fbDec.nMockStartScans := nScans;
END_METHOD

// #120: the stop of the mock axis ends at rest but never reports Done (a lost Done, or a stop that was never allowed)
METHOD SetStopWithoutDone
VAR_INPUT
	bHa		: BOOL;
	bDec	: BOOL;
END_VAR
fbHa.bMockNoStopDone := bHa;
fbDec.bMockNoStopDone := bDec;
END_METHOD

// the user offsets of the telescope under test (degrees; IAG50cm#17 telemetry tests)
METHOD SetOffsets
VAR_INPUT
	fHourAngle	: LREAL;
	fDeclination	: LREAL;
END_VAR
fbTel.HourAngleOffset := fHourAngle;
fbTel.DeclinationOffset := fDeclination;
END_METHOD

// the command input bStop of the telescope under test, as an ADS writer sets it (not the method)
METHOD SetStopInput
VAR_INPUT
	bValue	: BOOL;
END_VAR
fbTel.bStop := bValue;
END_METHOD

// the command input bPark of the telescope under test, as an ADS writer sets it (not the method)
METHOD SetParkInput
VAR_INPUT
	bValue	: BOOL;
END_VAR
fbTel.bPark := bValue;
END_METHOD

// the command input bPower of the telescope under test, as an ADS writer sets it (not the method)
METHOD SetPowerInput
VAR_INPUT
	bValue	: BOOL;
END_VAR
fbTel.bPower := bValue;
END_METHOD

// the command input bSlew of the telescope under test, as an ADS writer sets it (not the method)
METHOD SetSlewInput
VAR_INPUT
	bValue	: BOOL;
END_VAR
fbTel.bSlew := bValue;
END_METHOD

// the slew target fields an ADS writer sets before it raises bSlew
METHOD SetSlewTargetInput
VAR_INPUT
	fAzimuth	: LREAL;
	fAltitude	: LREAL;
END_VAR
fbTel.fAzimuth := fAzimuth;
fbTel.fElevation := fAltitude;
END_METHOD

// the command input bTrack of the telescope under test, as an ADS writer sets it (not the method)
METHOD SetTrackInput
VAR_INPUT
	bValue	: BOOL;
END_VAR
fbTel.bTrack := bValue;
END_METHOD

// sets the request latch bGoHomeActive of the telescope under test (an output, written through a pointer): a request left over from before

METHOD ForceGoHomeActive
pBool := ADR(fbTel.bGoHomeActive);

pBool^ := TRUE;
END_METHOD

// sets the request latch bSlewActive of the telescope under test (an output, written through a pointer): a request left over from before

METHOD ForceSlewActive
pBool := ADR(fbTel.bSlewActive);

pBool^ := TRUE;
END_METHOD

// the pointing-model safe altitude of the telescope under test (an input of the telescope; a goto target below it is refused)

METHOD SetSafeAltitude

VAR_INPUT

	fValue	: LREAL;

END_VAR
fbTel.fPointingSafeAltitude := fValue;
END_METHOD

// the E-stop input of the telescope under test (#14)
METHOD SetEstop
VAR_INPUT
	bValue	: BOOL;
END_VAR
fbTel.bEstopTriggered := bValue;
END_METHOD

METHOD InjectHaError
VAR_INPUT
	nId	: UDINT;
END_VAR
fbHa.InjectError(nId);
END_METHOD

METHOD InjectDecError
VAR_INPUT
	nId	: UDINT;
END_VAR
fbDec.InjectError(nId);
END_METHOD

END_FUNCTION_BLOCK

// ---- POUs/FB_RecordingComm.TcPOU
// I_Comm stub that records the Publish* calls of a test (parameter name, kind, value), for the telemetry characterization
// (IagTelemetry_Tests). Like FB_NullComm every call reports success. Recording is off until Start(), so the suites that
// do not look at the telemetry pay only the memory.
// Kinds: 1 LREAL, 2 INT (value as LREAL), 3 BOOL (0.0/1.0), 4 STRING (value not kept), 5 Publish (not kept).
FUNCTION_BLOCK FB_RecordingComm IMPLEMENTS BROTLib.I_Comm
VAR_OUTPUT
	nCount		: INT;			// records in aNames/aKinds/aValues (1..nCount)
	bOverflow	: BOOL;			// more than 160 calls: the last slot holds the newest call
	aNames		: ARRAY[1..160] OF STRING(80);
	aKinds		: ARRAY[1..160] OF INT;
	aValues		: ARRAY[1..160] OF LREAL;
END_VAR
VAR
	bRecording	: BOOL;
	sFilter		: STRING(80);
END_VAR

METHOD Publish : BOOL
VAR_INPUT
	domain			: STRING(255) := 'environment';
	location		: STRING(255) := 'roof';
	parameter		: STRING(255);
	value			: STRING(255);
END_VAR
VAR_OUTPUT
	published	: BOOL;
END_VAR
Record(sName := parameter, nKind := 5, fValue := 0.0);
Publish := TRUE;
published := TRUE;
END_METHOD

METHOD PublishLREAL : BOOL
VAR_INPUT
	domain			: STRING(255) := 'environment';
	location		: STRING(255) := 'roof';
	parameter		: STRING(255);
	value			: LREAL;
END_VAR
VAR_OUTPUT
	published	: BOOL;
END_VAR
Record(sName := parameter, nKind := 1, fValue := value);
PublishLREAL := TRUE;
published := TRUE;
END_METHOD

METHOD PublishINT : BOOL
VAR_INPUT
	domain			: STRING(255) := 'environment';
	location		: STRING(255) := 'roof';
	parameter		: STRING(255);
	value			: LINT;
END_VAR
VAR_OUTPUT
	published	: BOOL;
END_VAR
Record(sName := parameter, nKind := 2, fValue := LINT_TO_LREAL(value));
PublishINT := TRUE;
published := TRUE;
END_METHOD

METHOD PublishBOOL : BOOL
VAR_INPUT
	domain			: STRING(255) := 'environment';
	location		: STRING(255) := 'roof';
	parameter		: STRING(255);
	value			: BOOL;
END_VAR
VAR_OUTPUT
	published	: BOOL;
END_VAR
Record(sName := parameter, nKind := 3, fValue := SEL(value, 0.0, 1.0));
PublishBOOL := TRUE;
published := TRUE;
END_METHOD

METHOD PublishString : BOOL
VAR_INPUT
	domain			: STRING(255) := 'environment';
	location		: STRING(255) := 'roof';
	parameter		: STRING(255);
	value			: STRING(255);
END_VAR
VAR_OUTPUT
	published	: BOOL;
END_VAR
Record(sName := parameter, nKind := 4, fValue := 0.0);
PublishString := TRUE;
published := TRUE;
END_METHOD

METHOD PublishLog : BOOL
VAR_INPUT
	level		: STRING(255) := 'INFO';
	message		: STRING(255);
END_VAR
VAR_OUTPUT
	published	: BOOL;
END_VAR
PublishLog := TRUE;
published := TRUE;
END_METHOD

METHOD PRIVATE Record
VAR_INPUT
	sName	: STRING(255);
	nKind	: INT;
	fValue	: LREAL;
END_VAR
VAR
	nIndex	: INT;
END_VAR
IF NOT bRecording THEN
	RETURN;
END_IF
IF sFilter <> '' AND sFilter <> sName THEN
	RETURN;
END_IF
IF nCount >= 160 THEN
	// full: the last slot keeps the latest call, so a filtered recording still ends with the newest value
	bOverflow := TRUE;
	nIndex := 160;
ELSE
	nCount := nCount + 1;
	nIndex := nCount;
END_IF
aNames[nIndex] := sName;
aKinds[nIndex] := nKind;
aValues[nIndex] := fValue;
END_METHOD

// Clears the record and starts recording; sNameFilter <> '' records only calls with that parameter name.
METHOD Start
VAR_INPUT
	sNameFilter	: STRING(80);
END_VAR
VAR
	i	: INT;
END_VAR
FOR i := 1 TO 160 DO
	aNames[i] := '';
	aKinds[i] := 0;
	aValues[i] := 0.0;
END_FOR
nCount := 0;
bOverflow := FALSE;
sFilter := sNameFilter;
bRecording := TRUE;
END_METHOD

METHOD Stop
bRecording := FALSE;
END_METHOD

// first record with this parameter name, 0 if none
METHOD FindName : INT
VAR_INPUT
	sName	: STRING(80);
END_VAR
VAR
	i	: INT;
END_VAR
FindName := 0;
FOR i := 1 TO nCount DO
	IF aNames[i] = sName THEN
		FindName := i;
		RETURN;
	END_IF
END_FOR
END_METHOD

END_FUNCTION_BLOCK

// ---- POUs/F_Note.TcPOU
// Records a failed check in GVL_Diag.sFailures (see there). Called next to the TcUnit assertion, which does the actual test result.
FUNCTION F_Note : BOOL
VAR_INPUT
	bFailed	: BOOL;
	sText	: STRING(255);
END_VAR

IF bFailed AND LEN(GVL_Diag.sFailures) < 700 THEN
	GVL_Diag.sFailures := CONCAT(CONCAT(GVL_Diag.sFailures, sText), '; ');
END_IF
F_Note := bFailed;

END_FUNCTION

// ---- POUs/F_NoteNear.TcPOU
// TRUE (and a line in GVL_Diag.sFailures through F_Note) if fActual is not within fDelta of fExpected. NaN counts as failed.
FUNCTION F_NoteNear : BOOL
VAR_INPUT
	sText		: STRING(120);
	fExpected	: LREAL;
	fActual		: LREAL;
	fDelta		: LREAL;
END_VAR
VAR
	bNote		: BOOL;
END_VAR

F_NoteNear := NOT (ABS(fExpected - fActual) <= fDelta);
IF F_NoteNear THEN
	bNote := F_Note(bFailed := TRUE, sText := CONCAT(CONCAT(CONCAT(CONCAT(CONCAT(sText, ': expected '), LREAL_TO_STRING(fExpected)), ' +-'), LREAL_TO_STRING(fDelta)), CONCAT(', got ', LREAL_TO_STRING(fActual))));
END_IF

END_FUNCTION

// ---- POUs/IagResetUnderMotion_Tests.TcPOU
// Characterization of FB_TelescopeControl (IAG50cm) for a reset without and with an axis error, on mock axes (plan step 2,
// IAG50cmTests README). These tests pin what the code does today, with the line of the behaviour in a comment; they are not a
// specification. Every test owns a rig and runs over many PLC cycles (VAR_INST of the method, one Scan() per cycle). Failed checks
// are also noted in GVL_Diag.sFailures (printed by Run-Tests.ps1).
FUNCTION_BLOCK IagResetUnderMotion_Tests EXTENDS TcUnit.FB_TestSuite
VAR
END_VAR

Reset_Without_An_Error_Stops_The_Slew();
Reset_With_An_Error_Resets_The_Errored_Axis_And_Later_All_Axes();

// Command model step 3B.4: a reset without an error is a command to stop what moves: the slew latch is dropped and the moving axis gets one
// stop (abort stop). The hardware part stays gated: no axis is reset, no safety acknowledge is requested, the telescope stays online.
METHOD PRIVATE Reset_Without_An_Error_Stops_The_Slew
VAR_INST
	rig			: FB_IagRig;
	nStep		: INT;
	nCycles		: UINT;
	sTest		: STRING(80);
END_VAR
TEST('Reset_Without_An_Error_Stops_The_Slew');
sTest := 'Reset_Without_An_Error_Stops_The_Slew: ';
IF nStep >= 90 THEN
	RETURN;
END_IF
rig.Scan();
nCycles := nCycles + 1;
CASE nStep OF
0:	// wait for the clock, then power on
	IF rig.ClockValid THEN
		rig.fbTel.Init();
		nStep := 10;
		nCycles := 0;
	ELSIF nCycles > 2000 THEN
		AssertTrue(Condition := FALSE, Message := 'the astronomical clock never became valid');
		F_Note(bFailed := TRUE, sText := CONCAT(sTest, 'the astronomical clock never became valid'));
		nStep := 99;
		TEST_FINISHED();
	END_IF
10:	// online: slew
	IF rig.Online THEN
		rig.fbTel.Slew(fAzimuth := 180.0, fAltitude := 45.0);
		nStep := 20;
		nCycles := 0;
	ELSIF nCycles > 1500 THEN
		AssertTrue(Condition := FALSE, Message := 'the mock telescope did not reach READY_STATE 1.0');
		F_Note(bFailed := TRUE, sText := CONCAT(sTest, 'the mock telescope did not reach READY_STATE 1.0'));
		nStep := 99;
		TEST_FINISHED();
	END_IF
20:	// one axis is moving (the slew moves HA and Dec one after the other)
	IF rig.fbHa.MoveAxis OR rig.fbDec.MoveAxis THEN
		nStep := 30;
		nCycles := 0;
	ELSIF nCycles > 300 THEN
		AssertTrue(Condition := FALSE, Message := 'the slew did not start an axis move');
		F_Note(bFailed := TRUE, sText := CONCAT(sTest, 'the slew did not start an axis move'));
		nStep := 99;
		TEST_FINISHED();
	END_IF
30:	// let the move run for a few scans, then reset
	IF nCycles >= 5 THEN
		rig.fbTel.Reset();
		nStep := 40;
		nCycles := 0;
	END_IF
40:
	IF nCycles >= 10 THEN
		AssertFalse(Condition := rig.fbTel.bSlewActive, Message := 'the slew is dropped');
		F_Note(bFailed := (rig.fbTel.bSlewActive), sText := CONCAT(sTest, 'the slew is dropped'));
		AssertTrue(Condition := rig.fbHa.nResetEdges = 0 AND rig.fbDec.nResetEdges = 0, Message := 'no axis was reset');
		F_Note(bFailed := NOT (rig.fbHa.nResetEdges = 0 AND rig.fbDec.nResetEdges = 0), sText := CONCAT(sTest, 'no axis was reset'));
		AssertTrue(Condition := rig.fbHa.nStopEdges + rig.fbDec.nStopEdges = 1, Message := 'the moving axis got one stop');
		F_Note(bFailed := NOT (rig.fbHa.nStopEdges + rig.fbDec.nStopEdges = 1), sText := CONCAT(sTest, 'the moving axis got one stop'));
		AssertFalse(Condition := rig.fbTel.bSafetyAckRequest, Message := 'no safety acknowledge is requested');
		F_Note(bFailed := (rig.fbTel.bSafetyAckRequest), sText := CONCAT(sTest, 'no safety acknowledge is requested'));
		AssertTrue(Condition := rig.fbTel.ReadyState = 1.0, Message := 'the telescope stays online');
		F_Note(bFailed := NOT (rig.fbTel.ReadyState = 1.0), sText := CONCAT(sTest, 'the telescope stays online'));
		nStep := 99;
		TEST_FINISHED();
	END_IF
END_CASE
END_METHOD

// I:266-275, 1407 (#11, #55, #103): a reset with an error resets the axis that has the error and requests the safety acknowledge;
// 2.5 s later (bAxisResetAfterAck) a second pass resets every axis that is errored or not enabled. The error disabled both axes, so
// the second pass resets the errored one again and the other one for the first time.
METHOD PRIVATE Reset_With_An_Error_Resets_The_Errored_Axis_And_Later_All_Axes
VAR_INST
	rig			: FB_IagRig;
	nStep		: INT;
	nCycles		: UINT;
	sTest		: STRING(80);
END_VAR
TEST('Reset_With_An_Error_Resets_The_Errored_Axis_And_Later_All_Axes');
sTest := 'Reset_With_An_Error_Resets_The_Errored_Axis_And_Later_All_Axes: ';
IF nStep >= 90 THEN
	RETURN;
END_IF
rig.Scan();
nCycles := nCycles + 1;
CASE nStep OF
0:	// wait for the clock, then power on
	IF rig.ClockValid THEN
		rig.fbTel.Init();
		nStep := 10;
		nCycles := 0;
	ELSIF nCycles > 2000 THEN
		AssertTrue(Condition := FALSE, Message := 'the astronomical clock never became valid');
		F_Note(bFailed := TRUE, sText := CONCAT(sTest, 'the astronomical clock never became valid'));
		nStep := 99;
		TEST_FINISHED();
	END_IF
10:	// online: the hour angle reports an error
	IF rig.Online THEN
		rig.InjectHaError(16#4550);
		nStep := 20;
		nCycles := 0;
	ELSIF nCycles > 1500 THEN
		AssertTrue(Condition := FALSE, Message := 'the mock telescope did not reach READY_STATE 1.0');
		F_Note(bFailed := TRUE, sText := CONCAT(sTest, 'the mock telescope did not reach READY_STATE 1.0'));
		nStep := 99;
		TEST_FINISHED();
	END_IF
20:	// the error is there
	IF rig.fbTel.bError THEN
		rig.fbTel.Reset();
		nStep := 30;
		nCycles := 0;
	ELSIF nCycles > 60 THEN
		AssertTrue(Condition := FALSE, Message := 'the error was not reported');
		F_Note(bFailed := TRUE, sText := CONCAT(sTest, 'the error was not reported'));
		nStep := 99;
		TEST_FINISHED();
	END_IF
30:	// first pass
	IF nCycles = 5 THEN
		AssertFalse(Condition := rig.fbTel.bError, Message := 'the reset cleared the error');
		F_Note(bFailed := (rig.fbTel.bError), sText := CONCAT(sTest, 'the reset cleared the error'));
		AssertTrue(Condition := rig.fbHa.nResetEdges = 1 AND rig.fbDec.nResetEdges = 0, Message := 'the first pass resets only the errored axis');
		F_Note(bFailed := NOT (rig.fbHa.nResetEdges = 1 AND rig.fbDec.nResetEdges = 0), sText := CONCAT(sTest, 'the first pass resets only the errored axis'));
		AssertTrue(Condition := rig.fbTel.bSafetyAckRequest, Message := 'the reset requests the safety acknowledge');
		F_Note(bFailed := NOT (rig.fbTel.bSafetyAckRequest), sText := CONCAT(sTest, 'the reset requests the safety acknowledge'));
		nStep := 40;
		nCycles := 0;
	END_IF
40:	// second pass, 2.5 s later
	IF rig.fbHa.nResetEdges >= 2 AND nCycles > 5 THEN
		AssertTrue(Condition := rig.fbHa.nResetEdges = 2 AND rig.fbDec.nResetEdges = 1, Message := 'the second pass resets both axes, they are not enabled');
		F_Note(bFailed := NOT (rig.fbHa.nResetEdges = 2 AND rig.fbDec.nResetEdges = 1), sText := CONCAT(sTest, 'the second pass resets both axes, they are not enabled'));
		AssertFalse(Condition := rig.fbTel.bAxisResetAfterAck, Message := 'the second pass is over');
		F_Note(bFailed := (rig.fbTel.bAxisResetAfterAck), sText := CONCAT(sTest, 'the second pass is over'));
		nStep := 99;
		TEST_FINISHED();
	ELSIF nCycles > 800 THEN
		AssertTrue(Condition := FALSE, Message := 'the second reset pass never came');
		F_Note(bFailed := TRUE, sText := CONCAT(sTest, 'the second reset pass never came'));
		nStep := 99;
		TEST_FINISHED();
	END_IF
END_CASE
END_METHOD

END_FUNCTION_BLOCK

// ---- POUs/IagErrorPark_Tests.TcPOU
// Characterization of FB_TelescopeControl (IAG50cm) for an axis error and for a park during an error or with the axes off, on mock
// axes (plan step 2, IAG50cmTests README). These tests pin what the code does today, with the line of the behaviour in a comment;
// they are not a specification. Every test owns a rig and runs over many PLC cycles (VAR_INST of the method, one Scan() per
// cycle). Failed checks are also noted in GVL_Diag.sFailures (printed by Run-Tests.ps1).
FUNCTION_BLOCK IagErrorPark_Tests EXTENDS TcUnit.FB_TestSuite
VAR
END_VAR

Axis_Error_Starts_The_Park_Without_Moving_The_Mount();
Park_During_An_Error_Closes_The_Covers_And_Parks_The_Dome();
Park_With_The_Axes_Off_Does_Not_Move_The_Mount();
Error_Park_With_A_Stop_In_The_Same_Scan_Runs_After_Settle();

// BROTLib#25 step 4.4d (Tim 2026-11-09): an axis error drops every move command, disables both axes and, like MONETcommon#86, starts the
// park by itself: covers closed, dome parked, mount not moved, bIsParked not set. The telescope reports READY_STATE -1.0.
// (Before: IAG started no park on its own and the covers stayed as they were.)
METHOD PRIVATE Axis_Error_Starts_The_Park_Without_Moving_The_Mount
VAR_INST
	rig			: FB_IagRig;
	nStep		: INT;
	nCycles		: UINT;
	sTest		: STRING(80);
END_VAR
TEST('Axis_Error_Starts_The_Park_Without_Moving_The_Mount');
sTest := 'Axis_Error_Starts_The_Park_Without_Moving_The_Mount: ';
IF nStep >= 90 THEN
	RETURN;
END_IF
rig.Scan();
nCycles := nCycles + 1;
CASE nStep OF
0:	// wait for the clock, then power on
	IF rig.ClockValid THEN
		rig.fbTel.Init();
		nStep := 10;
		nCycles := 0;
	ELSIF nCycles > 2000 THEN
		AssertTrue(Condition := FALSE, Message := 'the astronomical clock never became valid');
		F_Note(bFailed := TRUE, sText := CONCAT(sTest, 'the astronomical clock never became valid'));
		nStep := 99;
		TEST_FINISHED();
	END_IF
10:	// online: the hour angle reports an error
	IF rig.Online THEN
		rig.InjectHaError(16#4550);
		nStep := 20;
		nCycles := 0;
	ELSIF nCycles > 1500 THEN
		AssertTrue(Condition := FALSE, Message := 'the mock telescope did not reach READY_STATE 1.0');
		F_Note(bFailed := TRUE, sText := CONCAT(sTest, 'the mock telescope did not reach READY_STATE 1.0'));
		nStep := 99;
		TEST_FINISHED();
	END_IF
20:
	IF nCycles >= 60 THEN
		AssertTrue(Condition := rig.fbTel.bError, Message := 'the error is reported');
		F_Note(bFailed := NOT (rig.fbTel.bError), sText := CONCAT(sTest, 'the error is reported'));
		AssertFalse(Condition := rig.fbHa.bEnable OR rig.fbDec.bEnable, Message := 'both axes are disabled');
		F_Note(bFailed := (rig.fbHa.bEnable OR rig.fbDec.bEnable), sText := CONCAT(sTest, 'both axes are disabled'));
		AssertTrue(Condition := rig.fbCovers.bClosed AND rig.fbCovers.nCloseCalls >= 1, Message := 'the error started the park: covers closed');
		F_Note(bFailed := NOT (rig.fbCovers.bClosed AND rig.fbCovers.nCloseCalls >= 1), sText := CONCAT(sTest, 'the error started the park: covers closed'));
		AssertTrue(Condition := rig.fbDome.nParkCalls >= 1, Message := 'the dome is parked');
		F_Note(bFailed := NOT (rig.fbDome.nParkCalls >= 1), sText := CONCAT(sTest, 'the dome is parked'));
		AssertFalse(Condition := rig.fbTel.bParkActive, Message := 'the park command is consumed');
		F_Note(bFailed := (rig.fbTel.bParkActive), sText := CONCAT(sTest, 'the park command is consumed'));
		AssertFalse(Condition := rig.fbHa.MoveAxis OR rig.fbDec.MoveAxis, Message := 'the mount was not moved');
		F_Note(bFailed := (rig.fbHa.MoveAxis OR rig.fbDec.MoveAxis), sText := CONCAT(sTest, 'the mount was not moved'));
		AssertFalse(Condition := rig.fbTel.bIsPowered, Message := 'the powered state is cleared by the error (#100)');
		F_Note(bFailed := rig.fbTel.bIsPowered, sText := CONCAT(sTest, 'the powered state is cleared by the error (#100)'));
		AssertTrue(Condition := rig.fbTel.ReadyState = -1.0, Message := 'READY_STATE is -1.0 (error)');
		F_Note(bFailed := NOT (rig.fbTel.ReadyState = -1.0), sText := CONCAT(sTest, 'READY_STATE is -1.0 (error)'));
		nStep := 99;
		TEST_FINISHED();
	END_IF
END_CASE
END_METHOD

// I:555-630: a park requested during an error does what is safe without the mount: the covers are closed, the dome is parked, the
// focus is disabled and the command is dropped. The mount is not moved and bIsParked is not set.
METHOD PRIVATE Park_During_An_Error_Closes_The_Covers_And_Parks_The_Dome
VAR_INST
	rig			: FB_IagRig;
	nStep		: INT;
	nCycles		: UINT;
	sTest		: STRING(80);
END_VAR
TEST('Park_During_An_Error_Closes_The_Covers_And_Parks_The_Dome');
sTest := 'Park_During_An_Error_Closes_The_Covers_And_Parks_The_Dome: ';
IF nStep >= 90 THEN
	RETURN;
END_IF
rig.Scan();
nCycles := nCycles + 1;
CASE nStep OF
0:	// wait for the clock, then power on
	IF rig.ClockValid THEN
		rig.fbTel.Init();
		nStep := 10;
		nCycles := 0;
	ELSIF nCycles > 2000 THEN
		AssertTrue(Condition := FALSE, Message := 'the astronomical clock never became valid');
		F_Note(bFailed := TRUE, sText := CONCAT(sTest, 'the astronomical clock never became valid'));
		nStep := 99;
		TEST_FINISHED();
	END_IF
10:	// online: the hour angle reports an error
	IF rig.Online THEN
		rig.InjectHaError(16#4550);
		nStep := 20;
		nCycles := 0;
	ELSIF nCycles > 1500 THEN
		AssertTrue(Condition := FALSE, Message := 'the mock telescope did not reach READY_STATE 1.0');
		F_Note(bFailed := TRUE, sText := CONCAT(sTest, 'the mock telescope did not reach READY_STATE 1.0'));
		nStep := 99;
		TEST_FINISHED();
	END_IF
20:	// the error is there: park
	IF rig.fbTel.bError THEN
		rig.fbTel.Park();
		nStep := 30;
		nCycles := 0;
	ELSIF nCycles > 60 THEN
		AssertTrue(Condition := FALSE, Message := 'the error was not reported');
		F_Note(bFailed := TRUE, sText := CONCAT(sTest, 'the error was not reported'));
		nStep := 99;
		TEST_FINISHED();
	END_IF
30:
	IF nCycles >= 30 THEN
		AssertTrue(Condition := rig.fbCovers.bClosed AND rig.fbCovers.nCloseCalls >= 1, Message := 'the covers are closed');
		F_Note(bFailed := NOT (rig.fbCovers.bClosed AND rig.fbCovers.nCloseCalls >= 1), sText := CONCAT(sTest, 'the covers are closed'));
		AssertTrue(Condition := rig.fbDome.nParkCalls >= 1, Message := 'the dome is parked');
		F_Note(bFailed := NOT (rig.fbDome.nParkCalls >= 1), sText := CONCAT(sTest, 'the dome is parked'));
		AssertFalse(Condition := rig.fbTel.bParkActive, Message := 'the park command is dropped');
		F_Note(bFailed := (rig.fbTel.bParkActive), sText := CONCAT(sTest, 'the park command is dropped'));
		AssertFalse(Condition := rig.fbTel.bIsParked, Message := 'the mount is not parked');
		F_Note(bFailed := (rig.fbTel.bIsParked), sText := CONCAT(sTest, 'the mount is not parked'));
		AssertFalse(Condition := rig.fbHa.MoveAxis OR rig.fbDec.MoveAxis, Message := 'the mount was not moved');
		F_Note(bFailed := (rig.fbHa.MoveAxis OR rig.fbDec.MoveAxis), sText := CONCAT(sTest, 'the mount was not moved'));
		AssertTrue(Condition := rig.fbTel.ReadyState = -1.0, Message := 'READY_STATE stays -1.0 (error)');
		F_Note(bFailed := NOT (rig.fbTel.ReadyState = -1.0), sText := CONCAT(sTest, 'READY_STATE stays -1.0 (error)'));
		nStep := 99;
		TEST_FINISHED();
	END_IF
END_CASE
END_METHOD

// I:555-600 (#54): a park on a telescope whose axes are off (never powered on) cannot drive the mount: the covers are closed and the
// dome parked, nothing moves. bIsParked is TRUE from the start (FB_TelescopeControl.bIsParked := TRUE) and the park leaves it.
METHOD PRIVATE Park_With_The_Axes_Off_Does_Not_Move_The_Mount
VAR_INST
	rig			: FB_IagRig;
	nStep		: INT;
	nCycles		: UINT;
	sTest		: STRING(80);
END_VAR
TEST('Park_With_The_Axes_Off_Does_Not_Move_The_Mount');
sTest := 'Park_With_The_Axes_Off_Does_Not_Move_The_Mount: ';
IF nStep >= 90 THEN
	RETURN;
END_IF
rig.Scan();
nCycles := nCycles + 1;
CASE nStep OF
0:	// wait for the clock
	IF rig.ClockValid THEN
		nStep := 10;
		nCycles := 0;
	ELSIF nCycles > 2000 THEN
		AssertTrue(Condition := FALSE, Message := 'the astronomical clock never became valid');
		F_Note(bFailed := TRUE, sText := CONCAT(sTest, 'the astronomical clock never became valid'));
		nStep := 99;
		TEST_FINISHED();
	END_IF
10:	// the axes are off: park
	rig.fbTel.Park();
	nStep := 20;
	nCycles := 0;
20:
	IF nCycles >= 30 THEN
		AssertTrue(Condition := rig.fbCovers.bClosed AND rig.fbCovers.nCloseCalls >= 1, Message := 'the covers are closed');
		F_Note(bFailed := NOT (rig.fbCovers.bClosed AND rig.fbCovers.nCloseCalls >= 1), sText := CONCAT(sTest, 'the covers are closed'));
		AssertTrue(Condition := rig.fbDome.nParkCalls >= 1, Message := 'the dome is parked');
		F_Note(bFailed := NOT (rig.fbDome.nParkCalls >= 1), sText := CONCAT(sTest, 'the dome is parked'));
		AssertFalse(Condition := rig.fbTel.bParkActive, Message := 'the park command is dropped');
		F_Note(bFailed := (rig.fbTel.bParkActive), sText := CONCAT(sTest, 'the park command is dropped'));
		AssertTrue(Condition := rig.fbTel.bIsParked, Message := 'bIsParked is still TRUE, as from the start: the park changes nothing');
		F_Note(bFailed := NOT (rig.fbTel.bIsParked), sText := CONCAT(sTest, 'bIsParked is still TRUE, as from the start: the park changes nothing'));
		AssertFalse(Condition := rig.fbHa.MoveAxis OR rig.fbDec.MoveAxis, Message := 'the mount was not moved');
		F_Note(bFailed := (rig.fbHa.MoveAxis OR rig.fbDec.MoveAxis), sText := CONCAT(sTest, 'the mount was not moved'));
		nStep := 99;
		TEST_FINISHED();
	END_IF
END_CASE
END_METHOD

// Characterization for the move of the error-park request (template body step S1.e): a stop in the scan of a new axis error queues the park behind it (bParkAfterStop); the park runs when the stop has settled. Written first, green before and after the move.
METHOD PRIVATE Error_Park_With_A_Stop_In_The_Same_Scan_Runs_After_Settle
VAR_INST
	rig			: FB_IagRig;
	nStep		: INT;
	nCycles		: UINT;
	sTest		: STRING(80);
END_VAR
TEST('Error_Park_With_A_Stop_In_The_Same_Scan_Runs_After_Settle');
sTest := 'Error_Park_With_A_Stop_In_The_Same_Scan_Runs_After_Settle: ';
IF nStep >= 90 THEN
	RETURN;
END_IF
rig.Scan();
nCycles := nCycles + 1;
CASE nStep OF
0:	// wait for the clock, then power on
	IF rig.ClockValid THEN
		rig.fbTel.Init();
		nStep := 10;
		nCycles := 0;
	ELSIF nCycles > 2000 THEN
		AssertTrue(Condition := FALSE, Message := 'the astronomical clock never became valid');
		F_Note(bFailed := TRUE, sText := CONCAT(sTest, 'the astronomical clock never became valid'));
		nStep := 99;
		TEST_FINISHED();
	END_IF
10:	// wait until the startup has finished (READY_STATE 1.0)
	IF rig.Online THEN
		rig.fbTel.Stop();
		rig.InjectHaError(16#4550);
		nStep := 20;
		nCycles := 0;
	ELSIF nCycles > 1500 THEN
		AssertTrue(Condition := FALSE, Message := 'the mock telescope did not reach READY_STATE 1.0');
		F_Note(bFailed := TRUE, sText := CONCAT(sTest, 'the mock telescope did not reach READY_STATE 1.0'));
		nStep := 99;
		TEST_FINISHED();
	END_IF
20:	// the error park is queued behind the stop and runs when the stop has settled
	IF nCycles >= 600 THEN
		AssertTrue(Condition := rig.fbTel.bError, Message := 'the error is reported');
		F_Note(bFailed := NOT (rig.fbTel.bError), sText := CONCAT(sTest, 'the error is reported'));
		AssertTrue(Condition := rig.fbCovers.bClosed AND rig.fbCovers.nCloseCalls >= 1, Message := 'the park ran after the stop: covers closed');
		F_Note(bFailed := NOT (rig.fbCovers.bClosed AND rig.fbCovers.nCloseCalls >= 1), sText := CONCAT(sTest, 'the park ran after the stop: covers closed'));
		AssertTrue(Condition := rig.fbDome.nParkCalls >= 1, Message := 'the dome is parked');
		F_Note(bFailed := NOT (rig.fbDome.nParkCalls >= 1), sText := CONCAT(sTest, 'the dome is parked'));
		AssertTrue(Condition := NOT rig.fbTel.bParkActive, Message := 'the park command is consumed');
		F_Note(bFailed := NOT (NOT rig.fbTel.bParkActive), sText := CONCAT(sTest, 'the park command is consumed'));
		AssertTrue(Condition := NOT rig.fbTel.bStopActive, Message := 'the stop is released');
		F_Note(bFailed := NOT (NOT rig.fbTel.bStopActive), sText := CONCAT(sTest, 'the stop is released'));
		nStep := 99;
		TEST_FINISHED();
	END_IF
END_CASE
END_METHOD

END_FUNCTION_BLOCK

// ---- POUs/IagTimeouts_Tests.TcPOU
// Characterization of the long timeouts of FB_TelescopeControl (IAG50cm) on mock axes, through the time seam (FB_TelescopeControl.nTimeDivisor,
// per rig; BROTLib FB_TimeoutTimer). Plan step 3 (decision 4). Failed checks are also noted in GVL_Diag.sFailures.
FUNCTION_BLOCK IagTimeouts_Tests EXTENDS TcUnit.FB_TestSuite
VAR
END_VAR

Slew_Times_Out_After_600_Seconds();
Idle_Telescope_Parks_After_12_Hours();

